(****************************************************************************************************<br>
© Syntegon Group.<br>
All rights reserved, also regarding any disposal, exploitation, reproduction, editing, distribution,<br>
as well as in the event of applications for industrial property rights.<br>
*****************************************************************************************************<br>
DESCRIPTION:<br>
A vision system's m_Configure describes housing, lens and the field of view as a frustum down to the working<br>
distance; a negative working distance gives a flat field of view at the lens.<br>
****************************************************************************************************)
METHOD PRIVATE m_VisionConfigure
VAR_INST
	fb_TempVision						: _FB_VisuVision;
	b_TempDone							: BOOL;	// the test ran
END_VAR
TEST('VisionConfigure');
IF b_TempDone THEN
	RETURN;
END_IF
b_TempDone := TRUE;

AssertTrue(Condition := fb_TempVision.m_Configure(vi_lr_FieldLength := 400, vi_lr_FieldWidth := 300,
	vi_lr_WorkingDistance := 800), Message := 'configured');
AssertEquals_UINT(Expected := 3, Actual := fb_TempVision.vo_Visu.stConfig.nBodyCount, Message := 'housing, lens, field of view');
AssertTrue(Condition := fb_TempVision.vo_Visu.stConfig.aBodies[2].eShape = E_VisuBodyShape.FRUSTUM,
	Message := 'field of view is a frustum');
AssertTrue(Condition := fb_TempVision.vo_Visu.stConfig.aBodies[2].eRole = E_VisuBodyRole.FIELD_OF_VIEW, Message := 'field of view role');
AssertEquals_LREAL(Expected := 800, Actual := fb_TempVision.vo_Visu.stConfig.aBodies[2].fHeight, Delta := 0.001,
	Message := 'field of view reaches the working distance');
AssertEquals_LREAL(Expected := -800, Actual := fb_TempVision.vo_Visu.stConfig.aBodies[2].stPose.fZ, Delta := 0.001,
	Message := 'field of view stands at the working distance below the lens');
AssertEquals_LREAL(Expected := 400, Actual := fb_TempVision.vo_Visu.stConfig.aBodies[2].fLength, Delta := 0.001,
	Message := 'field length at the bottom');

fb_TempVision.m_Configure(vi_lr_FieldLength := 400, vi_lr_FieldWidth := 300, vi_lr_WorkingDistance := -50);
AssertEquals_LREAL(Expected := 0, Actual := fb_TempVision.vo_Visu.stConfig.aBodies[2].fHeight, Delta := 0.001,
	Message := 'negative working distance: flat field of view');

TEST_FINISHED();
END_METHOD

END_FUNCTION_BLOCK

// ---- POUs/Tests/_FB_TestMachine.TcPOU
(****************************************************************************************************<br>
© Syntegon Group.<br>
All rights reserved, also regarding any disposal, exploitation, reproduction, editing, distribution,<br>
as well as in the event of applications for industrial property rights.<br>
*****************************************************************************************************<br>
DESCRIPTION:<br>
TcUnit test suite of _FB_VisuMachine: run state and simulation mode in the machine entry, machine messages set<br>
by their level, gone messages kept, and a full register making room with its oldest gone message.<br>
*****************************************************************************************************<br>
VERSION         ¦ DATE       ¦ NAME      ¦ CHANGE<br>
Syn_Visu 9.7.0  ¦ 2026-11-13 ¦ J.Willner ¦ Unit tests of the machine entry (protocol 22)<br>
****************************************************************************************************)
FUNCTION_BLOCK _FB_TestMachine EXTENDS TcUnit.FB_TestSuite
VAR
END_VAR

m_RunStateAndSimulation();
m_MessageRaisedAndCleared();
m_MessageIdZeroRefused();
m_FullRegisterMakesRoom();

(****************************************************************************************************<br>
© Syntegon Group.<br>
All rights reserved, also regarding any disposal, exploitation, reproduction, editing, distribution,<br>
as well as in the event of applications for industrial property rights.<br>
*****************************************************************************************************<br>
DESCRIPTION:<br>
A register full of active messages refuses a new one. Once some are gone, a new message takes the place of the<br>
oldest gone one (by its time): the others keep their order, the new one is last.<br>
****************************************************************************************************)
METHOD PRIVATE m_FullRegisterMakesRoom
VAR_INST
	fb_TempMachine						: _FB_VisuMachine;
	TempMachine							: ST_VisuMachine;
	b_TempDone							: BOOL;	// the test ran
END_VAR
VAR
	un_TempIndex						: UINT;
END_VAR
TEST('FullRegisterMakesRoom');
IF b_TempDone THEN
	RETURN;
END_IF
b_TempDone := TRUE;

fb_TempMachine.m_Register(vio_Machine := TempMachine);
FOR un_TempIndex := 1 TO VISU_GlobalConst_Param.VISU_un_MAX_MACHINE_MESSAGES DO
	fb_TempMachine.m_SetMessage(vi_udn_Id := un_TempIndex, vi_b_Active := TRUE,
		vi_e_Severity := E_VisuMessageSeverity.INFO, vi_str_Text := '', vi_udn_ComponentId := 0);
END_FOR
AssertEquals_UINT(Expected := VISU_GlobalConst_Param.VISU_un_MAX_MACHINE_MESSAGES, Actual := TempMachine.nMessageCount,
	Message := 'register full');
AssertFalse(Condition := fb_TempMachine.m_SetMessage(vi_udn_Id := 100, vi_b_Active := TRUE,
	vi_e_Severity := E_VisuMessageSeverity.INFO, vi_str_Text := '', vi_udn_ComponentId := 0),
	Message := 'full of active messages: a new one is refused');

(* Messages 3 and 5 go; 5 appeared earlier, so it is the oldest gone one. *)
fb_TempMachine.m_SetMessage(vi_udn_Id := 3, vi_b_Active := FALSE, vi_e_Severity := E_VisuMessageSeverity.INFO,
	vi_str_Text := '', vi_udn_ComponentId := 0);
fb_TempMachine.m_SetMessage(vi_udn_Id := 5, vi_b_Active := FALSE, vi_e_Severity := E_VisuMessageSeverity.INFO,
	vi_str_Text := '', vi_udn_ComponentId := 0);
TempMachine.aMessages[2].nTime := 2000;
TempMachine.aMessages[4].nTime := 1000;
AssertTrue(Condition := fb_TempMachine.m_SetMessage(vi_udn_Id := 100, vi_b_Active := TRUE,
	vi_e_Severity := E_VisuMessageSeverity.ERROR, vi_str_Text := 'New', vi_udn_ComponentId := 0),
	Message := 'with gone messages: a new one is listed');
AssertEquals_UINT(Expected := VISU_GlobalConst_Param.VISU_un_MAX_MACHINE_MESSAGES, Actual := TempMachine.nMessageCount,
	Message := 'still full');
AssertEquals_UDINT(Expected := 4, Actual := TempMachine.aMessages[3].nId, Message := 'message 4 before the gap');
AssertEquals_UDINT(Expected := 6, Actual := TempMachine.aMessages[4].nId, Message := 'message 5 left, 6 moved up');
AssertEquals_UDINT(Expected := 3, Actual := TempMachine.aMessages[2].nId, Message := 'message 3, gone later, stays');
AssertEquals_UDINT(Expected := 100, Actual := TempMachine.aMessages[VISU_GlobalConst_Param.VISU_un_MAX_MACHINE_MESSAGES - 1].nId,
	Message := 'the new message is last');
AssertTrue(Condition := TempMachine.aMessages[VISU_GlobalConst_Param.VISU_un_MAX_MACHINE_MESSAGES - 1].bActive,
	Message := 'the new message is active');

TEST_FINISHED();
END_METHOD

(****************************************************************************************************<br>
© Syntegon Group.<br>
All rights reserved, also regarding any disposal, exploitation, reproduction, editing, distribution,<br>
as well as in the event of applications for industrial property rights.<br>
*****************************************************************************************************<br>
DESCRIPTION:<br>
A message with id 0 is refused and not listed.<br>
****************************************************************************************************)
METHOD PRIVATE m_MessageIdZeroRefused
VAR_INST
	fb_TempMachine						: _FB_VisuMachine;
	TempMachine							: ST_VisuMachine;
	b_TempDone							: BOOL;	// the test ran
END_VAR
TEST('MessageIdZeroRefused');
IF b_TempDone THEN
	RETURN;
END_IF
b_TempDone := TRUE;

fb_TempMachine.m_Register(vio_Machine := TempMachine);
AssertFalse(Condition := fb_TempMachine.m_SetMessage(vi_udn_Id := 0, vi_b_Active := TRUE,
	vi_e_Severity := E_VisuMessageSeverity.ERROR, vi_str_Text := 'x', vi_udn_ComponentId := 0),
	Message := 'id 0 refused');
AssertEquals_UINT(Expected := 0, Actual := TempMachine.nMessageCount, Message := 'nothing listed');

TEST_FINISHED();
END_METHOD

(****************************************************************************************************<br>
© Syntegon Group.<br>
All rights reserved, also regarding any disposal, exploitation, reproduction, editing, distribution,<br>
as well as in the event of applications for industrial property rights.<br>
*****************************************************************************************************<br>
DESCRIPTION:<br>
A message set active is listed with its severity, text and component; set again it stays one entry and follows<br>
the inputs. Cleared it is gone but still listed; set active again it is the same entry, active once more. Clearing<br>
a message that was never listed lists nothing.<br>
****************************************************************************************************)
METHOD PRIVATE m_MessageRaisedAndCleared
VAR_INST
	fb_TempMachine						: _FB_VisuMachine;
	TempMachine							: ST_VisuMachine;
	b_TempDone							: BOOL;	// the test ran
END_VAR
TEST('MessageRaisedAndCleared');
IF b_TempDone THEN
	RETURN;
END_IF
b_TempDone := TRUE;

fb_TempMachine.m_Register(vio_Machine := TempMachine);
AssertTrue(Condition := fb_TempMachine.m_SetMessage(vi_udn_Id := 7, vi_b_Active := TRUE,
	vi_e_Severity := E_VisuMessageSeverity.WARNING, vi_str_Text := 'Reject bin almost full', vi_udn_ComponentId := 60),
	Message := 'a new message is listed');
AssertEquals_UINT(Expected := 1, Actual := TempMachine.nMessageCount, Message := 'one message');
AssertEquals_UDINT(Expected := 7, Actual := TempMachine.aMessages[0].nId, Message := 'its id');
AssertTrue(Condition := TempMachine.aMessages[0].bActive, Message := 'active');
AssertTrue(Condition := TempMachine.aMessages[0].eSeverity = E_VisuMessageSeverity.WARNING, Message := 'severity WARNING');
AssertEquals_STRING(Expected := 'Reject bin almost full', Actual := TempMachine.aMessages[0].sText, Message := 'its text');
AssertEquals_UDINT(Expected := 60, Actual := TempMachine.aMessages[0].nComponentId, Message := 'its component');

fb_TempMachine.m_SetMessage(vi_udn_Id := 7, vi_b_Active := TRUE, vi_e_Severity := E_VisuMessageSeverity.ERROR,
	vi_str_Text := 'Reject bin full', vi_udn_ComponentId := 60);
AssertEquals_UINT(Expected := 1, Actual := TempMachine.nMessageCount, Message := 'set again: still one message');
AssertTrue(Condition := TempMachine.aMessages[0].eSeverity = E_VisuMessageSeverity.ERROR, Message := 'severity follows');
AssertEquals_STRING(Expected := 'Reject bin full', Actual := TempMachine.aMessages[0].sText, Message := 'text follows');

fb_TempMachine.m_SetMessage(vi_udn_Id := 7, vi_b_Active := FALSE, vi_e_Severity := E_VisuMessageSeverity.ERROR,
	vi_str_Text := 'Reject bin full', vi_udn_ComponentId := 60);
AssertEquals_UINT(Expected := 1, Actual := TempMachine.nMessageCount, Message := 'cleared: still listed');
AssertFalse(Condition := TempMachine.aMessages[0].bActive, Message := 'cleared: gone');

fb_TempMachine.m_SetMessage(vi_udn_Id := 7, vi_b_Active := TRUE, vi_e_Severity := E_VisuMessageSeverity.ERROR,
	vi_str_Text := 'Reject bin full', vi_udn_ComponentId := 60);
AssertEquals_UINT(Expected := 1, Actual := TempMachine.nMessageCount, Message := 'raised again: the same entry');
AssertTrue(Condition := TempMachine.aMessages[0].bActive, Message := 'raised again: active');

AssertTrue(Condition := fb_TempMachine.m_SetMessage(vi_udn_Id := 8, vi_b_Active := FALSE,
	vi_e_Severity := E_VisuMessageSeverity.INFO, vi_str_Text := '', vi_udn_ComponentId := 0),
	Message := 'clearing an unlisted message succeeds');
AssertEquals_UINT(Expected := 1, Actual := TempMachine.nMessageCount, Message := '... and lists nothing');

TEST_FINISHED();
END_METHOD

(****************************************************************************************************<br>
© Syntegon Group.<br>
All rights reserved, also regarding any disposal, exploitation, reproduction, editing, distribution,<br>
as well as in the event of applications for industrial property rights.<br>
*****************************************************************************************************<br>
DESCRIPTION:<br>
Before m_Register the methods write nothing; after it the run state, its text and simulation mode are in the<br>
machine entry.<br>
****************************************************************************************************)
METHOD PRIVATE m_RunStateAndSimulation
VAR_INST
	fb_TempMachine						: _FB_VisuMachine;
	TempMachine							: ST_VisuMachine;
	b_TempDone							: BOOL;	// the test ran
END_VAR
TEST('RunStateAndSimulation');
IF b_TempDone THEN
	RETURN;
END_IF
b_TempDone := TRUE;

AssertFalse(Condition := fb_TempMachine.m_SetRunState(vi_e_RunState := E_VisuRunState.RUNNING, vi_str_Text := ''),
	Message := 'm_SetRunState before m_Register: FALSE');
AssertFalse(Condition := fb_TempMachine.m_SetMessage(vi_udn_Id := 1, vi_b_Active := TRUE,
	vi_e_Severity := E_VisuMessageSeverity.ERROR, vi_str_Text := 'x', vi_udn_ComponentId := 0),
	Message := 'm_SetMessage before m_Register: FALSE');

AssertTrue(Condition := fb_TempMachine.m_Register(vio_Machine := TempMachine), Message := 'm_Register');
AssertTrue(Condition := fb_TempMachine.m_SetRunState(vi_e_RunState := E_VisuRunState.FAULT, vi_str_Text := 'Vacuum lost'),
	Message := 'm_SetRunState after m_Register');
AssertTrue(Condition := fb_TempMachine.m_SetSimulation(vi_b_Simulation := TRUE), Message := 'm_SetSimulation');
AssertTrue(Condition := TempMachine.eRunState = E_VisuRunState.FAULT, Message := 'run state FAULT');
AssertEquals_STRING(Expected := 'Vacuum lost', Actual := TempMachine.sRunStateText, Message := 'run state text');
AssertTrue(Condition := TempMachine.bSimulation, Message := 'simulation mode');
AssertEquals_UINT(Expected := 0, Actual := TempMachine.nMessageCount, Message := 'no messages');

TEST_FINISHED();
END_METHOD

END_FUNCTION_BLOCK

// ---- POUs/Tests/_FB_TestConfigComponent.TcPOU
(****************************************************************************************************<br>
© Syntegon Group.<br>
All rights reserved, also regarding any disposal, exploitation, reproduction, editing, distribution,<br>
as well as in the event of applications for industrial property rights.<br>
*****************************************************************************************************<br>
DESCRIPTION:<br>
TcUnit test suite of SynConfig._FB_ConfigComponent: registration in the config manifest (m_Register, m_Id), the<br>
symbol path of vo_Config taken from the instance path, and the protocol and library version reported to the<br>
gateway.<br>
*****************************************************************************************************<br>
VERSION         ¦ DATE       ¦ NAME      ¦ CHANGE<br>
Syn_Config 2.0.0 ¦ 2026-11-11 ¦ J.Willner ¦ Unit tests<br>
****************************************************************************************************)
FUNCTION_BLOCK _FB_TestConfigComponent EXTENDS TcUnit.FB_TestSuite
VAR
	fb_PathConveyorParam				: SynConfig._FB_ConfigConveyor;	// declared here so that its instance path is known
END_VAR

m_RegisterAddsEntry();
m_RegisterIsIdempotent();
m_RegisterRejectsIdZero();
m_RegisterRejectsUsedId();
m_RegisterRejectsFullManifest();
m_RegisterSymbolPath();
m_VersionMatchesConstant();

(****************************************************************************************************<br>
© Syntegon Group.<br>
All rights reserved, also regarding any disposal, exploitation, reproduction, editing, distribution,<br>
as well as in the event of applications for industrial property rights.<br>
*****************************************************************************************************<br>
DESCRIPTION:<br>
m_Register adds an entry with the id and type of the parametrised component, gives the id through m_Id and<br>
reports the running library's protocol and library version in the manifest.<br>
****************************************************************************************************)
METHOD PRIVATE m_RegisterAddsEntry
VAR_INST
	fb_TempParam						: SynConfig._FB_ConfigDelta;
	TempManifest						: SynConfig.ST_ConfigManifest;
	b_TempDone							: BOOL;	// the test ran
END_VAR
TEST('ConfigRegisterAddsEntry');
IF b_TempDone THEN
	RETURN;
END_IF
b_TempDone := TRUE;

AssertEquals_UDINT(Expected := 0, Actual := fb_TempParam.m_Id(), Message := 'not registered: id 0');
AssertTrue(Condition := fb_TempParam.m_Register(vio_Manifest := TempManifest, vi_udn_Id := 10), Message := 'registered');
AssertEquals_UINT(Expected := 1, Actual := TempManifest.nCount, Message := 'one entry');
AssertEquals_UDINT(Expected := 10, Actual := TempManifest.aEntries[0].nId, Message := 'entry has the component id');
AssertTrue(Condition := TempManifest.aEntries[0].eType = E_VisuComponentType.DELTA, Message := 'entry has the component type');
AssertEquals_UDINT(Expected := 10, Actual := fb_TempParam.m_Id(), Message := 'm_Id gives the id');
AssertEquals_UINT(Expected := SynConfig.CONFIG_GlobalConst.CONFIG_un_PROTOCOL_VERSION, Actual := TempManifest.nProtocolVersion,
	Message := 'config protocol version reported');
AssertEquals_STRING(Expected := SynConfig.CONFIG_GlobalConst.CONFIG_str_LIBRARY_VERSION, Actual := TempManifest.sLibraryVersion,
	Message := 'library version reported');

TEST_FINISHED();
END_METHOD

(****************************************************************************************************<br>
© Syntegon Group.<br>
All rights reserved, also regarding any disposal, exploitation, reproduction, editing, distribution,<br>
as well as in the event of applications for industrial property rights.<br>
*****************************************************************************************************<br>
DESCRIPTION:<br>
m_Register is called every cycle: registering again with the same id succeeds without a second entry.<br>
****************************************************************************************************)
METHOD PRIVATE m_RegisterIsIdempotent
VAR_INST
	fb_TempParam						: SynConfig._FB_ConfigConveyor;
	TempManifest						: SynConfig.ST_ConfigManifest;
	b_TempDone							: BOOL;	// the test ran
END_VAR
TEST('ConfigRegisterIsIdempotent');
IF b_TempDone THEN
	RETURN;
END_IF
b_TempDone := TRUE;

AssertTrue(Condition := fb_TempParam.m_Register(vio_Manifest := TempManifest, vi_udn_Id := 1), Message := 'first call');
AssertTrue(Condition := fb_TempParam.m_Register(vio_Manifest := TempManifest, vi_udn_Id := 1), Message := 'second call');
AssertEquals_UINT(Expected := 1, Actual := TempManifest.nCount, Message := 'still one entry');

TEST_FINISHED();
END_METHOD

(****************************************************************************************************<br>
© Syntegon Group.<br>
All rights reserved, also regarding any disposal, exploitation, reproduction, editing, distribution,<br>
as well as in the event of applications for industrial property rights.<br>
*****************************************************************************************************<br>
DESCRIPTION:<br>
The config manifest takes CONFIG_un_MAX_MANIFEST_ENTRIES entries; a new id beyond them is refused.<br>
****************************************************************************************************)
METHOD PRIVATE m_RegisterRejectsFullManifest
VAR_INST
	fb_TempParam						: SynConfig._FB_ConfigConveyor;
	TempManifest						: SynConfig.ST_ConfigManifest;
	b_TempDone							: BOOL;	// the test ran
END_VAR
VAR
	un_TempEntry						: UINT;
END_VAR
TEST('ConfigRegisterRejectsFullManifest');
IF b_TempDone THEN
	RETURN;
END_IF
b_TempDone := TRUE;

(* Other parameter FBs have filled the manifest. *)
FOR un_TempEntry := 0 TO SynConfig.CONFIG_GlobalConst_Param.CONFIG_un_MAX_MANIFEST_ENTRIES - 1 DO
	TempManifest.aEntries[un_TempEntry].nId := UINT_TO_UDINT(un_TempEntry + 1);
	TempManifest.aEntries[un_TempEntry].eType := E_VisuComponentType.CONVEYOR;
	TempManifest.aEntries[un_TempEntry].sPath := 'P_Line.fb_Param.vo_Config';
END_FOR
TempManifest.nCount := SynConfig.CONFIG_GlobalConst_Param.CONFIG_un_MAX_MANIFEST_ENTRIES;

AssertFalse(Condition := fb_TempParam.m_Register(vio_Manifest := TempManifest, vi_udn_Id := 999), Message := 'full manifest refuses');
AssertEquals_UINT(Expected := SynConfig.CONFIG_GlobalConst_Param.CONFIG_un_MAX_MANIFEST_ENTRIES, Actual := TempManifest.nCount,
	Message := 'entry count at the limit');

TEST_FINISHED();
END_METHOD

(****************************************************************************************************<br>
© Syntegon Group.<br>
All rights reserved, also regarding any disposal, exploitation, reproduction, editing, distribution,<br>
as well as in the event of applications for industrial property rights.<br>
*****************************************************************************************************<br>
DESCRIPTION:<br>
Id 0 is no component (an unregistered Syn_Visu FB's m_Id): m_Register refuses it and adds nothing.<br>
****************************************************************************************************)
METHOD PRIVATE m_RegisterRejectsIdZero
VAR_INST
	fb_TempParam						: SynConfig._FB_ConfigConveyor;
	TempManifest						: SynConfig.ST_ConfigManifest;
	b_TempDone							: BOOL;	// the test ran
END_VAR
TEST('ConfigRegisterRejectsIdZero');
IF b_TempDone THEN
	RETURN;
END_IF
b_TempDone := TRUE;

AssertFalse(Condition := fb_TempParam.m_Register(vio_Manifest := TempManifest, vi_udn_Id := 0), Message := 'id 0 refused');
AssertEquals_UINT(Expected := 0, Actual := TempManifest.nCount, Message := 'no entry');
AssertEquals_UDINT(Expected := 0, Actual := fb_TempParam.m_Id(), Message := 'still not registered');

TEST_FINISHED();
END_METHOD

(****************************************************************************************************<br>
© Syntegon Group.<br>
All rights reserved, also regarding any disposal, exploitation, reproduction, editing, distribution,<br>
as well as in the event of applications for industrial property rights.<br>
*****************************************************************************************************<br>
DESCRIPTION:<br>
One parameter FB per component: an id already registered by another FB is refused, whether that FB has another<br>
type or the same type at another symbol path.<br>
****************************************************************************************************)
METHOD PRIVATE m_RegisterRejectsUsedId
VAR_INST
	fb_TempConveyorParam				: SynConfig._FB_ConfigConveyor;
	fb_TempOtherConveyorParam			: SynConfig._FB_ConfigConveyor;
	fb_TempDeltaParam					: SynConfig._FB_ConfigDelta;
	TempManifest						: SynConfig.ST_ConfigManifest;
	b_TempDone							: BOOL;	// the test ran
END_VAR
TEST('ConfigRegisterRejectsUsedId');
IF b_TempDone THEN
	RETURN;
END_IF
b_TempDone := TRUE;

AssertTrue(Condition := fb_TempConveyorParam.m_Register(vio_Manifest := TempManifest, vi_udn_Id := 3), Message := 'first FB registered');
AssertFalse(Condition := fb_TempDeltaParam.m_Register(vio_Manifest := TempManifest, vi_udn_Id := 3),
	Message := 'another type with the same id refused');
AssertFalse(Condition := fb_TempOtherConveyorParam.m_Register(vio_Manifest := TempManifest, vi_udn_Id := 3),
	Message := 'the same type at another path refused');
AssertEquals_UINT(Expected := 1, Actual := TempManifest.nCount, Message := 'still one entry');
AssertEquals_UDINT(Expected := 0, Actual := fb_TempDeltaParam.m_Id(), Message := 'refused FB not registered');

TEST_FINISHED();
END_METHOD

(****************************************************************************************************<br>
© Syntegon Group.<br>
All rights reserved, also regarding any disposal, exploitation, reproduction, editing, distribution,<br>
as well as in the event of applications for industrial property rights.<br>
*****************************************************************************************************<br>
DESCRIPTION:<br>
The manifest entry's symbol path is the instance path without TwinCAT project and PLC project, plus<br>
'.vo_Config': the path the gateway reads and writes over ADS.<br>
****************************************************************************************************)
METHOD PRIVATE m_RegisterSymbolPath
VAR_INST
	TempManifest						: SynConfig.ST_ConfigManifest;
	b_TempDone							: BOOL;	// the test ran
END_VAR
TEST('ConfigRegisterSymbolPath');
IF b_TempDone THEN
	RETURN;
END_IF
b_TempDone := TRUE;

fb_PathConveyorParam.m_Register(vio_Manifest := TempManifest, vi_udn_Id := 1);
AssertEquals_STRING(Expected := 'P_TestRun.fb_TestConfigComponent.fb_PathConveyorParam.vo_Config',
	Actual := TempManifest.aEntries[0].sPath, Message := 'symbol path of vo_Config without TwinCAT and PLC project');

TEST_FINISHED();
END_METHOD

(****************************************************************************************************<br>
© Syntegon Group.<br>
All rights reserved, also regarding any disposal, exploitation, reproduction, editing, distribution,<br>
as well as in the event of applications for industrial property rights.<br>
*****************************************************************************************************<br>
DESCRIPTION:<br>
_FC_GetVersionSynConfig and CONFIG_str_LIBRARY_VERSION name the same version: both are bumped together.<br>
****************************************************************************************************)
METHOD PRIVATE m_VersionMatchesConstant
VAR_INST
	b_TempDone							: BOOL;	// the test ran
END_VAR
VAR
	str_TempVersion						: STRING(31);	// major.minor.revision from _FC_GetVersionSynConfig
END_VAR
TEST('ConfigVersionMatchesConstant');
IF b_TempDone THEN
	RETURN;
END_IF
b_TempDone := TRUE;

str_TempVersion := CONCAT(UINT_TO_STRING(SynConfig._FC_GetVersionSynConfig(vi_n_VersionElement := 1)), '.');
str_TempVersion := CONCAT(str_TempVersion, UINT_TO_STRING(SynConfig._FC_GetVersionSynConfig(vi_n_VersionElement := 2)));
str_TempVersion := CONCAT(str_TempVersion, '.');
str_TempVersion := CONCAT(str_TempVersion, UINT_TO_STRING(SynConfig._FC_GetVersionSynConfig(vi_n_VersionElement := 3)));
AssertEquals_STRING(Expected := SynConfig.CONFIG_GlobalConst.CONFIG_str_LIBRARY_VERSION, Actual := str_TempVersion,
	Message := '_FC_GetVersionSynConfig matches CONFIG_str_LIBRARY_VERSION');
AssertEquals_UINT(Expected := 16#FFFF, Actual := SynConfig._FC_GetVersionSynConfig(vi_n_VersionElement := 4),
	Message := 'unknown version element gives 16#FFFF');

TEST_FINISHED();
END_METHOD

END_FUNCTION_BLOCK

// ---- POUs/Tests/_FB_TestConfigStaging.TcPOU
(****************************************************************************************************<br>
© Syntegon Group.<br>
All rights reserved, also regarding any disposal, exploitation, reproduction, editing, distribution,<br>
as well as in the event of applications for industrial property rights.<br>
*****************************************************************************************************<br>
DESCRIPTION:<br>
TcUnit test suite of a parameter FB's m_Cycle (ADR 0017), on SynConfig._FB_ConfigConveyor: the program values<br>
while no set is active, a staged set taken over, waiting while the application does not allow it, rejected on<br>
another active version or when invalid, and a reset back to the program values. The tests write vo_Config's<br>
stStaging and stStaged as the gateway does over ADS.<br>
*****************************************************************************************************<br>
VERSION         ¦ DATE       ¦ NAME      ¦ CHANGE<br>
Syn_Config 2.0.0 ¦ 2026-11-11 ¦ J.Willner ¦ Unit tests<br>
Syn_Config 2.3.0 ¦ 2026-11-14 ¦ J.Willner ¦ The lifecycle of every parameter FB type<br>
****************************************************************************************************)
FUNCTION_BLOCK _FB_TestConfigStaging EXTENDS TcUnit.FB_TestSuite

m_ProgramValuesWithoutSet();
m_StagedSetTakenOver();
m_StagedSetWaitsUntilAllowed();
m_StagedSetOnOtherVersionRejected();
m_ResetReturnsToProgramValues();
m_InvalidProductTypesRejected();
m_EveryTypeRunsTheLifecycle();

(****************************************************************************************************<br>
© Syntegon Group.<br>
All rights reserved, also regarding any disposal, exploitation, reproduction, editing, distribution,<br>
as well as in the event of applications for industrial property rights.<br>
*****************************************************************************************************<br>
DESCRIPTION:<br>
Every parameter FB type runs the same staging lifecycle as the conveyor: a set staged on version 0 is taken over<br>
as version 1, a set staged on version 0 again is rejected (version 1 is active), and a reset returns to the<br>
program values under version 0. The machine FB's recipe has its own suite (_FB_TestConfigMachine).<br>
****************************************************************************************************)
METHOD PRIVATE m_EveryTypeRunsTheLifecycle
VAR_INST
	fb_TempDelta						: SynConfig._FB_ConfigDelta;
	TempDeltaDefault					: SynConfig.ST_ConfigDeltaParam;
	TempDeltaStaged						: SynConfig.ST_ConfigDeltaParam;
	TempDeltaSet						: SynConfig.ST_ConfigDeltaSet;
	fb_TempGantry						: SynConfig._FB_ConfigXtsGantry;
	TempGantryDefault					: SynConfig.ST_ConfigXtsGantryParam;
	TempGantryStaged					: SynConfig.ST_ConfigXtsGantryParam;
	TempGantrySet						: SynConfig.ST_ConfigXtsGantrySet;
	fb_TempLoop							: SynConfig._FB_ConfigXtsLoop;
	TempLoopDefault						: SynConfig.ST_ConfigXtsLoopParam;
	TempLoopStaged						: SynConfig.ST_ConfigXtsLoopParam;
	TempLoopSet							: SynConfig.ST_ConfigXtsLoopSet;
	fb_TempCartesian					: SynConfig._FB_ConfigCartesian;
	TempCartesianDefault				: SynConfig.ST_ConfigCartesianParam;
	TempCartesianStaged					: SynConfig.ST_ConfigCartesianParam;
	TempCartesianSet					: SynConfig.ST_ConfigCartesianSet;
	fb_TempVision						: SynConfig._FB_ConfigVision;
	TempVisionDefault					: SynConfig.ST_ConfigBodyComponentParam;
	TempVisionStaged					: SynConfig.ST_ConfigBodyComponentParam;
	TempVisionSet						: SynConfig.ST_ConfigBodyComponentSet;
	b_TempDone							: BOOL;	// the test ran
END_VAR
VAR
	b_TempChanged						: ARRAY[1..5, 1..3] OF BOOL;	// per type and step: m_Cycle's result
	e_TempResult						: ARRAY[1..5, 1..3] OF SynConfig.E_ConfigResult;	// per type and step: stStatus.eResult
	udn_TempVersion						: ARRAY[1..5, 1..3] OF UDINT;	// [-] per type and step: stStatus.nActiveVersion
	lr_TempX							: ARRAY[1..5, 1..3] OF LREAL;	// [mm] per type and step: X of the effective pose
	TempPose							: ST_VisuPose;
	un_TempStep							: UINT;	// [-] 1 = take-over, 2 = stale version, 3 = reset
	un_TempType							: UINT;
	p_TempDelta							: POINTER TO SynConfig.ST_ConfigDeltaParam;
	p_TempGantry						: POINTER TO SynConfig.ST_ConfigXtsGantryParam;
	p_TempLoop							: POINTER TO SynConfig.ST_ConfigXtsLoopParam;
	p_TempCartesian						: POINTER TO SynConfig.ST_ConfigCartesianParam;
	p_TempVision						: POINTER TO SynConfig.ST_ConfigBodyComponentParam;
END_VAR
VAR CONSTANT
	str_TYPE_NAMES						: ARRAY[1..5] OF STRING(20) := ['Delta', 'XTS gantry', 'XTS loop', 'Cartesian', 'Vision'];
END_VAR
TEST('ConfigEveryTypeRunsTheLifecycle');
IF b_TempDone THEN
	RETURN;
END_IF
b_TempDone := TRUE;


(****************************************************************************************************
THREE STEPS PER TYPE: TAKE-OVER, STALE VERSION, RESET
****************************************************************************************************)
(* Delta *)
TempDeltaDefault.stPose.fX := 100;
TempDeltaStaged.stPose.fX := 250;
p_TempDelta := ADR(fb_TempDelta.vo_Config.stStaged);
FOR un_TempStep := 1 TO 3 DO
	p_TempDelta^ := TempDeltaStaged;
	_FC_TestConfigStage(vi_p_Staging := ADR(fb_TempDelta.vo_Config.stStaging), vi_udn_BaseVersion := 0,
		vi_udn_StageId := UINT_TO_UDINT(un_TempStep), vi_b_Reset := un_TempStep = 3);
	b_TempChanged[1, un_TempStep] := fb_TempDelta.m_Cycle(vio_Default := TempDeltaDefault, vio_Set := TempDeltaSet,
		vi_b_ApplyAllowed := TRUE);
	e_TempResult[1, un_TempStep] := fb_TempDelta.vo_Config.stStatus.eResult;
	udn_TempVersion[1, un_TempStep] := fb_TempDelta.vo_Config.stStatus.nActiveVersion;
	TempPose := fb_TempDelta.m_Pose();
	lr_TempX[1, un_TempStep] := TempPose.fX;
END_FOR

(* XTS gantry: a track needs a module *)
TempGantryDefault.stPose.fX := 100;
TempGantryStaged.stPose.fX := 250;
TempGantryStaged.nModuleCount := 1;
TempGantryStaged.aModules[0].fLength := 250;
p_TempGantry := ADR(fb_TempGantry.vo_Config.stStaged);
FOR un_TempStep := 1 TO 3 DO
	p_TempGantry^ := TempGantryStaged;
	_FC_TestConfigStage(vi_p_Staging := ADR(fb_TempGantry.vo_Config.stStaging), vi_udn_BaseVersion := 0,
		vi_udn_StageId := UINT_TO_UDINT(un_TempStep), vi_b_Reset := un_TempStep = 3);
	b_TempChanged[2, un_TempStep] := fb_TempGantry.m_Cycle(vio_Default := TempGantryDefault, vio_Set := TempGantrySet,
		vi_b_ApplyAllowed := TRUE);
	e_TempResult[2, un_TempStep] := fb_TempGantry.vo_Config.stStatus.eResult;
	udn_TempVersion[2, un_TempStep] := fb_TempGantry.vo_Config.stStatus.nActiveVersion;
	TempPose := fb_TempGantry.m_Pose();
	lr_TempX[2, un_TempStep] := TempPose.fX;
END_FOR

(* XTS loop: a track needs a module *)
TempLoopDefault.stPose.fX := 100;
TempLoopStaged.stPose.fX := 250;
TempLoopStaged.nModuleCount := 1;
TempLoopStaged.aModules[0].fLength := 250;
p_TempLoop := ADR(fb_TempLoop.vo_Config.stStaged);
FOR un_TempStep := 1 TO 3 DO
	p_TempLoop^ := TempLoopStaged;
	_FC_TestConfigStage(vi_p_Staging := ADR(fb_TempLoop.vo_Config.stStaging), vi_udn_BaseVersion := 0,
		vi_udn_StageId := UINT_TO_UDINT(un_TempStep), vi_b_Reset := un_TempStep = 3);
	b_TempChanged[3, un_TempStep] := fb_TempLoop.m_Cycle(vio_Default := TempLoopDefault, vio_Set := TempLoopSet,
		vi_b_ApplyAllowed := TRUE);
	e_TempResult[3, un_TempStep] := fb_TempLoop.vo_Config.stStatus.eResult;
	udn_TempVersion[3, un_TempStep] := fb_TempLoop.vo_Config.stStatus.nActiveVersion;
	TempPose := fb_TempLoop.m_Pose();
	lr_TempX[3, un_TempStep] := TempPose.fX;
END_FOR

(* Cartesian *)
TempCartesianDefault.stPose.fX := 100;
TempCartesianStaged.stPose.fX := 250;
p_TempCartesian := ADR(fb_TempCartesian.vo_Config.stStaged);
FOR un_TempStep := 1 TO 3 DO
	p_TempCartesian^ := TempCartesianStaged;
	_FC_TestConfigStage(vi_p_Staging := ADR(fb_TempCartesian.vo_Config.stStaging), vi_udn_BaseVersion := 0,
		vi_udn_StageId := UINT_TO_UDINT(un_TempStep), vi_b_Reset := un_TempStep = 3);
	b_TempChanged[4, un_TempStep] := fb_TempCartesian.m_Cycle(vio_Default := TempCartesianDefault,
		vio_Set := TempCartesianSet, vi_b_ApplyAllowed := TRUE);
	e_TempResult[4, un_TempStep] := fb_TempCartesian.vo_Config.stStatus.eResult;
	udn_TempVersion[4, un_TempStep] := fb_TempCartesian.vo_Config.stStatus.nActiveVersion;
	TempPose := fb_TempCartesian.m_Pose();
	lr_TempX[4, un_TempStep] := TempPose.fX;
END_FOR

(* Vision system, for the body components *)
TempVisionDefault.stPose.fX := 100;
TempVisionStaged.stPose.fX := 250;
p_TempVision := ADR(fb_TempVision.vo_Config.stStaged);
FOR un_TempStep := 1 TO 3 DO
	p_TempVision^ := TempVisionStaged;
	_FC_TestConfigStage(vi_p_Staging := ADR(fb_TempVision.vo_Config.stStaging), vi_udn_BaseVersion := 0,
		vi_udn_StageId := UINT_TO_UDINT(un_TempStep), vi_b_Reset := un_TempStep = 3);
	b_TempChanged[5, un_TempStep] := fb_TempVision.m_Cycle(vio_Default := TempVisionDefault, vio_Set := TempVisionSet,
		vi_b_ApplyAllowed := TRUE);
	e_TempResult[5, un_TempStep] := fb_TempVision.vo_Config.stStatus.eResult;
	udn_TempVersion[5, un_TempStep] := fb_TempVision.vo_Config.stStatus.nActiveVersion;
	TempPose := fb_TempVision.m_Pose();
	lr_TempX[5, un_TempStep] := TempPose.fX;
END_FOR


(****************************************************************************************************
THE SAME RESULTS FOR EVERY TYPE
****************************************************************************************************)
FOR un_TempType := 1 TO 5 DO
	AssertTrue(Condition := b_TempChanged[un_TempType, 1], Message := CONCAT(str_TYPE_NAMES[un_TempType], ': taken over'));
	AssertEquals_UDINT(Expected := 1, Actual := udn_TempVersion[un_TempType, 1],
		Message := CONCAT(str_TYPE_NAMES[un_TempType], ': version 1 active'));
	AssertEquals_LREAL(Expected := 250, Actual := lr_TempX[un_TempType, 1], Delta := 0.001,
		Message := CONCAT(str_TYPE_NAMES[un_TempType], ': staged pose effective'));
	AssertFalse(Condition := b_TempChanged[un_TempType, 2],
		Message := CONCAT(str_TYPE_NAMES[un_TempType], ': stale version not taken over'));
	AssertTrue(Condition := e_TempResult[un_TempType, 2] = SynConfig.E_ConfigResult.REJECTED,
		Message := CONCAT(str_TYPE_NAMES[un_TempType], ': stale version rejected'));
	AssertEquals_UDINT(Expected := 1, Actual := udn_TempVersion[un_TempType, 2],
		Message := CONCAT(str_TYPE_NAMES[un_TempType], ': version 1 stays'));
	AssertTrue(Condition := b_TempChanged[un_TempType, 3], Message := CONCAT(str_TYPE_NAMES[un_TempType], ': reset'));
	AssertEquals_UDINT(Expected := 0, Actual := udn_TempVersion[un_TempType, 3],
		Message := CONCAT(str_TYPE_NAMES[un_TempType], ': version 0 after the reset'));
	AssertEquals_LREAL(Expected := 100, Actual := lr_TempX[un_TempType, 3], Delta := 0.001,
		Message := CONCAT(str_TYPE_NAMES[un_TempType], ': program pose again'));
END_FOR

TEST_FINISHED();
END_METHOD

(****************************************************************************************************<br>
© Syntegon Group.<br>
All rights reserved, also regarding any disposal, exploitation, reproduction, editing, distribution,<br>
as well as in the event of applications for industrial property rights.<br>
*****************************************************************************************************<br>
DESCRIPTION:<br>
A conveyor set is rejected with the reason when a product type has no number, a number is used twice or there<br>
are more product types than the list holds; the active set stays as it was.<br>
****************************************************************************************************)
METHOD PRIVATE m_InvalidProductTypesRejected
VAR_INST
	fb_TempParam						: SynConfig._FB_ConfigConveyor;
	TempDefault							: SynConfig.ST_ConfigConveyorParam;
	TempSet								: SynConfig.ST_ConfigConveyorSet;
	b_TempDone							: BOOL;	// the test ran
END_VAR
VAR
	TempStaged							: SynConfig.ST_ConfigConveyorParam;
END_VAR
TEST('ConfigInvalidProductTypesRejected');
IF b_TempDone THEN
	RETURN;
END_IF
b_TempDone := TRUE;

TempDefault := m_ValidSet(vi_lr_X := 100);

(* A product type without a number. *)
TempStaged := m_ValidSet(vi_lr_X := 250);
TempStaged.aProductTypes[1].nId := 0;
m_Stage(vio_Param := fb_TempParam, vio_Staged := TempStaged, vi_udn_BaseVersion := 0, vi_udn_StageId := 1);
AssertFalse(Condition := fb_TempParam.m_Cycle(vio_Default := TempDefault, vio_Set := TempSet, vi_b_ApplyAllowed := TRUE),
	Message := 'type without a number: not taken over');
AssertTrue(Condition := fb_TempParam.vo_Config.stStatus.eResult = SynConfig.E_ConfigResult.REJECTED, Message := 'rejected');
AssertEquals_STRING(Expected := 'A product type without a number', Actual := fb_TempParam.vo_Config.stStatus.sMessage,
	Message := 'reason: no number');

(* A number used twice. *)
TempStaged := m_ValidSet(vi_lr_X := 250);
TempStaged.aProductTypes[0].nId := 3;
TempStaged.aProductTypes[1].nId := 3;
m_Stage(vio_Param := fb_TempParam, vio_Staged := TempStaged, vi_udn_BaseVersion := 0, vi_udn_StageId := 2);
AssertFalse(Condition := fb_TempParam.m_Cycle(vio_Default := TempDefault, vio_Set := TempSet, vi_b_ApplyAllowed := TRUE),
	Message := 'number twice: not taken over');
AssertEquals_STRING(Expected := 'Product type 3 is defined twice', Actual := fb_TempParam.vo_Config.stStatus.sMessage,
	Message := 'reason: defined twice');

(* More product types than the list holds. *)
TempStaged := m_ValidSet(vi_lr_X := 250);
TempStaged.nProductTypeCount := VISU_GlobalConst_Param.VISU_un_MAX_PRODUCT_TYPES + 1;
m_Stage(vio_Param := fb_TempParam, vio_Staged := TempStaged, vi_udn_BaseVersion := 0, vi_udn_StageId := 3);
AssertFalse(Condition := fb_TempParam.m_Cycle(vio_Default := TempDefault, vio_Set := TempSet, vi_b_ApplyAllowed := TRUE),
	Message := 'too many types: not taken over');
AssertEquals_STRING(Expected := CONCAT('More than ', CONCAT(UINT_TO_STRING(VISU_GlobalConst_Param.VISU_un_MAX_PRODUCT_TYPES),
	' product types')), Actual := fb_TempParam.vo_Config.stStatus.sMessage, Message := 'reason: too many');
AssertEquals_UDINT(Expected := 3, Actual := fb_TempParam.vo_Config.stStatus.nHandledStageId, Message := 'last stage id handled');

AssertFalse(Condition := TempSet.bValid, Message := 'still no active set');
AssertEquals_LREAL(Expected := 100, Actual := fb_TempParam.vo_Config.stActive.stPose.fX, Delta := 0.001,
	Message := 'program values still effective');

TEST_FINISHED();
END_METHOD

(****************************************************************************************************<br>
© Syntegon Group.<br>
All rights reserved, also regarding any disposal, exploitation, reproduction, editing, distribution,<br>
as well as in the event of applications for industrial property rights.<br>
*****************************************************************************************************<br>
DESCRIPTION:<br>
Without an active set the program values are effective, under version 0, and nothing has been handled.<br>
****************************************************************************************************)
METHOD PRIVATE m_ProgramValuesWithoutSet
VAR_INST
	fb_TempParam						: SynConfig._FB_ConfigConveyor;
	TempDefault							: SynConfig.ST_ConfigConveyorParam;
	TempSet								: SynConfig.ST_ConfigConveyorSet;
	b_TempDone							: BOOL;	// the test ran
END_VAR
VAR
	TempPose							: ST_VisuPose;
END_VAR
TEST('ConfigProgramValuesWithoutSet');
IF b_TempDone THEN
	RETURN;
END_IF
b_TempDone := TRUE;

TempDefault := m_ValidSet(vi_lr_X := 100);
AssertFalse(Condition := fb_TempParam.m_Cycle(vio_Default := TempDefault, vio_Set := TempSet, vi_b_ApplyAllowed := TRUE),
	Message := 'nothing staged: no change');
TempPose := fb_TempParam.m_Pose();
AssertEquals_LREAL(Expected := 100, Actual := TempPose.fX, Delta := 0.001, Message := 'program pose effective');
AssertEquals_UINT(Expected := 2, Actual := fb_TempParam.vo_Config.stActive.nProductTypeCount, Message := 'program product types effective');
AssertEquals_UDINT(Expected := 0, Actual := fb_TempParam.vo_Config.stStatus.nActiveVersion, Message := 'version 0: program values');
AssertTrue(Condition := fb_TempParam.vo_Config.stStatus.eResult = SynConfig.E_ConfigResult.NONE, Message := 'nothing handled');

TEST_FINISHED();
END_METHOD

(****************************************************************************************************<br>
© Syntegon Group.<br>
All rights reserved, also regarding any disposal, exploitation, reproduction, editing, distribution,<br>
as well as in the event of applications for industrial property rights.<br>
*****************************************************************************************************<br>
DESCRIPTION:<br>
A reset makes the active set invalid at once (also while a take-over is not allowed): the program values apply<br>
under version 0. Versions never repeat: the next set taken over gets version 2, not 1.<br>
****************************************************************************************************)
METHOD PRIVATE m_ResetReturnsToProgramValues
VAR_INST
	fb_TempParam						: SynConfig._FB_ConfigConveyor;
	TempDefault							: SynConfig.ST_ConfigConveyorParam;
	TempSet								: SynConfig.ST_ConfigConveyorSet;
	b_TempDone							: BOOL;	// the test ran
END_VAR
VAR
	TempStaged							: SynConfig.ST_ConfigConveyorParam;
END_VAR
TEST('ConfigResetReturnsToProgramValues');
IF b_TempDone THEN
	RETURN;
END_IF
b_TempDone := TRUE;

TempDefault := m_ValidSet(vi_lr_X := 100);
TempStaged := m_ValidSet(vi_lr_X := 250);
m_Stage(vio_Param := fb_TempParam, vio_Staged := TempStaged, vi_udn_BaseVersion := 0, vi_udn_StageId := 1);
fb_TempParam.m_Cycle(vio_Default := TempDefault, vio_Set := TempSet, vi_b_ApplyAllowed := TRUE);
AssertEquals_UDINT(Expected := 1, Actual := fb_TempParam.vo_Config.stStatus.nActiveVersion, Message := 'version 1 active');

_FC_TestConfigStage(vi_p_Staging := ADR(fb_TempParam.vo_Config.stStaging), vi_udn_BaseVersion := 1, vi_udn_StageId := 2,
	vi_b_Reset := TRUE);
AssertTrue(Condition := fb_TempParam.m_Cycle(vio_Default := TempDefault, vio_Set := TempSet, vi_b_ApplyAllowed := FALSE),
	Message := 'reset handled, even while not allowed');
AssertFalse(Condition := TempSet.bValid, Message := 'active set invalid');
AssertEquals_UDINT(Expected := 0, Actual := fb_TempParam.vo_Config.stStatus.nActiveVersion, Message := 'version 0');
AssertEquals_LREAL(Expected := 100, Actual := fb_TempParam.vo_Config.stActive.stPose.fX, Delta := 0.001,
	Message := 'program values effective again');
AssertTrue(Condition := fb_TempParam.vo_Config.stStatus.eResult = SynConfig.E_ConfigResult.APPLIED, Message := 'reset applied');
AssertEquals_UDINT(Expected := 2, Actual := fb_TempParam.vo_Config.stStatus.nHandledStageId, Message := 'stage id handled');
AssertFalse(Condition := fb_TempParam.vo_Config.stStaging.bReset, Message := 'reset flag cleared');

m_Stage(vio_Param := fb_TempParam, vio_Staged := TempStaged, vi_udn_BaseVersion := 0, vi_udn_StageId := 3);
fb_TempParam.m_Cycle(vio_Default := TempDefault, vio_Set := TempSet, vi_b_ApplyAllowed := TRUE);
AssertEquals_UDINT(Expected := 2, Actual := fb_TempParam.vo_Config.stStatus.nActiveVersion, Message := 'next set gets version 2');

TEST_FINISHED();
END_METHOD

(****************************************************************************************************<br>
© Syntegon Group.<br>
All rights reserved, also regarding any disposal, exploitation, reproduction, editing, distribution,<br>
as well as in the event of applications for industrial property rights.<br>
*****************************************************************************************************<br>
DESCRIPTION:<br>
Stages a set on a conveyor's parameter FB as the gateway does: the set into vo_Config.stStaged, then stStaging<br>
(_FC_TestConfigStage). The FB handles it in its next m_Cycle.<br>
****************************************************************************************************)
METHOD PRIVATE m_Stage : BOOL
VAR_IN_OUT
	vio_Param							: SynConfig._FB_ConfigConveyor;	// the parameter FB under test
END_VAR
VAR_IN_OUT CONSTANT
	vio_Staged							: SynConfig.ST_ConfigConveyorParam;	// the set to stage
END_VAR
VAR_INPUT
	vi_udn_BaseVersion					: UDINT;	// [-] active version the set is based on
	vi_udn_StageId						: UDINT;	// [-] the gateway's id of this staging
END_VAR
VAR
	p_TempStaged						: POINTER TO SynConfig.ST_ConfigConveyorParam;
END_VAR
p_TempStaged := ADR(vio_Param.vo_Config.stStaged);
p_TempStaged^ := vio_Staged;
m_Stage := _FC_TestConfigStage(vi_p_Staging := ADR(vio_Param.vo_Config.stStaging), vi_udn_BaseVersion := vi_udn_BaseVersion,
	vi_udn_StageId := vi_udn_StageId, vi_b_Reset := FALSE);
END_METHOD

(****************************************************************************************************<br>
© Syntegon Group.<br>
All rights reserved, also regarding any disposal, exploitation, reproduction, editing, distribution,<br>
as well as in the event of applications for industrial property rights.<br>
*****************************************************************************************************<br>
DESCRIPTION:<br>
A set staged on another version than the active one is rejected with the reason, even while a take-over is<br>
allowed: someone else changed the set since the configurator read it.<br>
****************************************************************************************************)
METHOD PRIVATE m_StagedSetOnOtherVersionRejected
VAR_INST
	fb_TempParam						: SynConfig._FB_ConfigConveyor;
	TempDefault							: SynConfig.ST_ConfigConveyorParam;
	TempSet								: SynConfig.ST_ConfigConveyorSet;
	b_TempDone							: BOOL;	// the test ran
END_VAR
VAR
	TempStaged							: SynConfig.ST_ConfigConveyorParam;
END_VAR
TEST('ConfigStagedSetOnOtherVersionRejected');
IF b_TempDone THEN
	RETURN;
END_IF
b_TempDone := TRUE;

TempDefault := m_ValidSet(vi_lr_X := 100);
TempStaged := m_ValidSet(vi_lr_X := 250);
m_Stage(vio_Param := fb_TempParam, vio_Staged := TempStaged, vi_udn_BaseVersion := 5, vi_udn_StageId := 9);

AssertFalse(Condition := fb_TempParam.m_Cycle(vio_Default := TempDefault, vio_Set := TempSet, vi_b_ApplyAllowed := TRUE),
	Message := 'not taken over');
AssertTrue(Condition := fb_TempParam.vo_Config.stStatus.eResult = SynConfig.E_ConfigResult.REJECTED, Message := 'rejected');
AssertEquals_STRING(Expected := 'Based on version 5, but version 0 is active', Actual := fb_TempParam.vo_Config.stStatus.sMessage,
	Message := 'the reason');
AssertEquals_UDINT(Expected := 9, Actual := fb_TempParam.vo_Config.stStatus.nHandledStageId, Message := 'stage id handled');
AssertFalse(Condition := fb_TempParam.vo_Config.stStaging.bStaged, Message := 'staged flag cleared');
AssertFalse(Condition := TempSet.bValid, Message := 'no active set');

TEST_FINISHED();
END_METHOD

(****************************************************************************************************<br>
© Syntegon Group.<br>
All rights reserved, also regarding any disposal, exploitation, reproduction, editing, distribution,<br>
as well as in the event of applications for industrial property rights.<br>
*****************************************************************************************************<br>
DESCRIPTION:<br>
A set staged on the active version is taken over while the application allows it: it becomes the active set<br>
under version 1 and the effective values, the status names the stage id as applied and the flags are cleared.<br>
****************************************************************************************************)
METHOD PRIVATE m_StagedSetTakenOver
VAR_INST
	fb_TempParam						: SynConfig._FB_ConfigConveyor;
	TempDefault							: SynConfig.ST_ConfigConveyorParam;
	TempSet								: SynConfig.ST_ConfigConveyorSet;
	b_TempDone							: BOOL;	// the test ran
END_VAR
VAR
	TempPose							: ST_VisuPose;
	TempStaged							: SynConfig.ST_ConfigConveyorParam;
END_VAR
TEST('ConfigStagedSetTakenOver');
IF b_TempDone THEN
	RETURN;
END_IF
b_TempDone := TRUE;

TempDefault := m_ValidSet(vi_lr_X := 100);
TempStaged := m_ValidSet(vi_lr_X := 250);
m_Stage(vio_Param := fb_TempParam, vio_Staged := TempStaged, vi_udn_BaseVersion := 0, vi_udn_StageId := 7);

AssertTrue(Condition := fb_TempParam.m_Cycle(vio_Default := TempDefault, vio_Set := TempSet, vi_b_ApplyAllowed := TRUE),
	Message := 'set taken over');
AssertTrue(Condition := TempSet.bValid, Message := 'active set valid');
AssertEquals_UDINT(Expected := 1, Actual := TempSet.nVersion, Message := 'first version');
AssertEquals_UDINT(Expected := 1, Actual := fb_TempParam.vo_Config.stStatus.nActiveVersion, Message := 'status names the version');
AssertEquals_UDINT(Expected := 7, Actual := fb_TempParam.vo_Config.stStatus.nHandledStageId, Message := 'stage id handled');
AssertTrue(Condition := fb_TempParam.vo_Config.stStatus.eResult = SynConfig.E_ConfigResult.APPLIED, Message := 'applied');
AssertEquals_STRING(Expected := '', Actual := fb_TempParam.vo_Config.stStatus.sMessage, Message := 'no message');
AssertFalse(Condition := fb_TempParam.vo_Config.stStaging.bStaged, Message := 'staged flag cleared');
TempPose := fb_TempParam.m_Pose();
AssertEquals_LREAL(Expected := 250, Actual := TempPose.fX, Delta := 0.001, Message := 'staged pose effective');

AssertFalse(Condition := fb_TempParam.m_Cycle(vio_Default := TempDefault, vio_Set := TempSet, vi_b_ApplyAllowed := TRUE),
	Message := 'next cycle: no change');
AssertEquals_UDINT(Expected := 1, Actual := fb_TempParam.vo_Config.stStatus.nActiveVersion, Message := 'still version 1');

TEST_FINISHED();
END_METHOD

(****************************************************************************************************<br>
© Syntegon Group.<br>
All rights reserved, also regarding any disposal, exploitation, reproduction, editing, distribution,<br>
as well as in the event of applications for industrial property rights.<br>
*****************************************************************************************************<br>
DESCRIPTION:<br>
While the application does not allow a take-over the staged set waits (PENDING, still staged, the program values<br>
stay effective); it is taken over in the first cycle that allows it.<br>
****************************************************************************************************)
METHOD PRIVATE m_StagedSetWaitsUntilAllowed
VAR_INST
	fb_TempParam						: SynConfig._FB_ConfigConveyor;
	TempDefault							: SynConfig.ST_ConfigConveyorParam;
	TempSet								: SynConfig.ST_ConfigConveyorSet;
	b_TempDone							: BOOL;	// the test ran
END_VAR
VAR
	TempStaged							: SynConfig.ST_ConfigConveyorParam;
END_VAR
TEST('ConfigStagedSetWaitsUntilAllowed');
IF b_TempDone THEN
	RETURN;
END_IF
b_TempDone := TRUE;

TempDefault := m_ValidSet(vi_lr_X := 100);
TempStaged := m_ValidSet(vi_lr_X := 250);
m_Stage(vio_Param := fb_TempParam, vio_Staged := TempStaged, vi_udn_BaseVersion := 0, vi_udn_StageId := 3);

AssertFalse(Condition := fb_TempParam.m_Cycle(vio_Default := TempDefault, vio_Set := TempSet, vi_b_ApplyAllowed := FALSE),
	Message := 'not allowed: not taken over');
AssertTrue(Condition := fb_TempParam.vo_Config.stStatus.eResult = SynConfig.E_ConfigResult.PENDING, Message := 'pending');
AssertTrue(Condition := fb_TempParam.vo_Config.stStaging.bStaged, Message := 'still staged');
AssertFalse(Condition := TempSet.bValid, Message := 'no active set yet');
AssertEquals_LREAL(Expected := 100, Actual := fb_TempParam.vo_Config.stActive.stPose.fX, Delta := 0.001,
	Message := 'program values still effective');

AssertTrue(Condition := fb_TempParam.m_Cycle(vio_Default := TempDefault, vio_Set := TempSet, vi_b_ApplyAllowed := TRUE),
	Message := 'allowed: taken over');
AssertTrue(Condition := fb_TempParam.vo_Config.stStatus.eResult = SynConfig.E_ConfigResult.APPLIED, Message := 'applied');
AssertEquals_UDINT(Expected := 3, Actual := fb_TempParam.vo_Config.stStatus.nHandledStageId, Message := 'stage id handled');

TEST_FINISHED();
END_METHOD

(****************************************************************************************************<br>
© Syntegon Group.<br>
All rights reserved, also regarding any disposal, exploitation, reproduction, editing, distribution,<br>
as well as in the event of applications for industrial property rights.<br>
*****************************************************************************************************<br>
DESCRIPTION:<br>
A conveyor parameter set that can be taken over: the pose at X = vi_lr_X and two product types (1 and 2).<br>
****************************************************************************************************)
METHOD PRIVATE m_ValidSet : SynConfig.ST_ConfigConveyorParam
VAR_INPUT
	vi_lr_X								: LREAL;	// [mm] X of the pose, to tell sets apart
END_VAR
m_ValidSet.stPose.fX := vi_lr_X;
m_ValidSet.stOriginShift.fX := 50;
m_ValidSet.nProductTypeCount := 2;
m_ValidSet.aProductTypes[0].nId := 1;
m_ValidSet.aProductTypes[0].fLength := 120;
m_ValidSet.aProductTypes[0].fWidth := 80;
m_ValidSet.aProductTypes[0].fHeight := 40;
m_ValidSet.aProductTypes[0].eShape := E_VisuProductShape.BOX;
m_ValidSet.aProductTypes[1].nId := 2;
m_ValidSet.aProductTypes[1].fLength := 66;
m_ValidSet.aProductTypes[1].fWidth := 66;
m_ValidSet.aProductTypes[1].fHeight := 120;
m_ValidSet.aProductTypes[1].eShape := E_VisuProductShape.CYLINDER;
END_METHOD

END_FUNCTION_BLOCK

// ---- POUs/Tests/_FC_TestConfigStage.TcPOU
(****************************************************************************************************<br>
© Syntegon Group.<br>
All rights reserved, also regarding any disposal, exploitation, reproduction, editing, distribution,<br>
as well as in the event of applications for industrial property rights.<br>
*****************************************************************************************************<br>
DESCRIPTION:<br>
Writes a parameter FB's stStaging as the gateway does over ADS (docs/config-contract.md): the version the set is<br>
based on, a stage id, and bStaged (a set, written to stStaged before) or bReset last. ST cannot assign to an FB's<br>
output, so the tests pass the address of vo_Config.stStaging, as ADS writes into the PLC's memory.<br>
*****************************************************************************************************<br>
OUTPUT VALUES:<br>
FALSE for a null pointer.<br>
*****************************************************************************************************<br>
VERSION         ¦ DATE       ¦ NAME      ¦ CHANGE<br>
Syn_Config 2.0.0 ¦ 2026-11-11 ¦ J.Willner ¦ Unit tests<br>
****************************************************************************************************)
FUNCTION _FC_TestConfigStage : BOOL
VAR_INPUT
	vi_p_Staging						: POINTER TO SynConfig.ST_ConfigStaging;	// ADR(fb_Param.vo_Config.stStaging)
	vi_udn_BaseVersion					: UDINT;	// [-] active version the set is based on
	vi_udn_StageId						: UDINT;	// [-] the gateway's id of this staging
	vi_b_Reset							: BOOL;	// [-] TRUE: a reset instead of a staged set
END_VAR

_FC_TestConfigStage := vi_p_Staging <> 0;
IF NOT _FC_TestConfigStage THEN
	RETURN;
END_IF
vi_p_Staging^.bStaged := FALSE;
vi_p_Staging^.nBaseVersion := vi_udn_BaseVersion;
vi_p_Staging^.nStageId := vi_udn_StageId;
vi_p_Staging^.bReset := vi_b_Reset;
vi_p_Staging^.bStaged := NOT vi_b_Reset;

END_FUNCTION

// ---- POUs/Tests/_FB_TestConfigRobot.TcPOU
(****************************************************************************************************<br>
© Syntegon Group.<br>
All rights reserved, also regarding any disposal, exploitation, reproduction, editing, distribution,<br>
as well as in the event of applications for industrial property rights.<br>
*****************************************************************************************************<br>
DESCRIPTION:<br>
TcUnit test suite of the robots' parameter FBs (SynConfig._FB_ConfigDelta, _FB_ConfigXtsGantry,<br>
_FB_ConfigXtsLoop, _FB_ConfigCartesian): which staged sets are rejected and why (zones, gripper fingers, track<br>
modules), and m_PassOn handing the effective values on to the robot's Syn_Visu FB, its config version changing<br>
only when a value does, its lists shrinking with the set.<br>
*****************************************************************************************************<br>
VERSION         ¦ DATE       ¦ NAME      ¦ CHANGE<br>
Syn_Config 2.0.0 ¦ 2026-11-11 ¦ J.Willner ¦ Unit tests<br>
****************************************************************************************************)
FUNCTION_BLOCK _FB_TestConfigRobot EXTENDS TcUnit.FB_TestSuite

m_DeltaRejectsInvalidZonesAndFingers();
m_XtsTracksRejectInvalidModules();
m_CartesianTakesOverFingers();
m_DeltaPassOn();
m_DeltaPassOnShrinksLists();
m_XtsGantryPassOnModules();

(****************************************************************************************************<br>
© Syntegon Group.<br>
All rights reserved, also regarding any disposal, exploitation, reproduction, editing, distribution,<br>
as well as in the event of applications for industrial property rights.<br>
*****************************************************************************************************<br>
DESCRIPTION:<br>
A Cartesian robot's set takes its gripper fingers over with their offsets on the flange (ADR 0018); a finger<br>
without a height is rejected.<br>
****************************************************************************************************)
METHOD PRIVATE m_CartesianTakesOverFingers
VAR_INST
	fb_TempParam						: SynConfig._FB_ConfigCartesian;
	TempDefault							: SynConfig.ST_ConfigCartesianParam;
	TempSet								: SynConfig.ST_ConfigCartesianSet;
	b_TempDone							: BOOL;	// the test ran
END_VAR
VAR
	TempStaged							: SynConfig.ST_ConfigCartesianParam;
	p_TempStaged						: POINTER TO SynConfig.ST_ConfigCartesianParam;
END_VAR
TEST('ConfigCartesianTakesOverFingers');
IF b_TempDone THEN
	RETURN;
END_IF
b_TempDone := TRUE;

p_TempStaged := ADR(fb_TempParam.vo_Config.stStaged);
TempStaged.nFingerCount := 2;
TempStaged.aFingers[0].fDiameter := 30;
TempStaged.aFingers[0].fHeight := 60;
TempStaged.aFingers[1].fDiameter := 30;
TempStaged.aFingers[1].fHeight := 0;
TempStaged.aFingers[1].stOffset.fY := -45;
TempStaged.aFingers[1].stOffset.fRz := 90;

p_TempStaged^ := TempStaged;
_FC_TestConfigStage(vi_p_Staging := ADR(fb_TempParam.vo_Config.stStaging), vi_udn_BaseVersion := 0, vi_udn_StageId := 1,
	vi_b_Reset := FALSE);
AssertFalse(Condition := fb_TempParam.m_Cycle(vio_Default := TempDefault, vio_Set := TempSet, vi_b_ApplyAllowed := TRUE),
	Message := 'finger without a height: not taken over');
AssertEquals_STRING(Expected := 'Finger 2 has no diameter or height', Actual := fb_TempParam.vo_Config.stStatus.sMessage,
	Message := 'reason');

TempStaged.aFingers[1].fHeight := 60;
p_TempStaged^ := TempStaged;
_FC_TestConfigStage(vi_p_Staging := ADR(fb_TempParam.vo_Config.stStaging), vi_udn_BaseVersion := 0, vi_udn_StageId := 2,
	vi_b_Reset := FALSE);
AssertTrue(Condition := fb_TempParam.m_Cycle(vio_Default := TempDefault, vio_Set := TempSet, vi_b_ApplyAllowed := TRUE),
	Message := 'valid fingers taken over');
AssertEquals_UINT(Expected := 2, Actual := fb_TempParam.vo_Config.stActive.nFingerCount, Message := 'two fingers effective');
AssertEquals_LREAL(Expected := -45, Actual := fb_TempParam.vo_Config.stActive.aFingers[1].stOffset.fY, Delta := 0.001,
	Message := 'offset Y kept');
AssertEquals_LREAL(Expected := 90, Actual := fb_TempParam.vo_Config.stActive.aFingers[1].stOffset.fRz, Delta := 0.001,
	Message := 'offset rotation kept');

TEST_FINISHED();
END_METHOD

(****************************************************************************************************<br>
© Syntegon Group.<br>
All rights reserved, also regarding any disposal, exploitation, reproduction, editing, distribution,<br>
as well as in the event of applications for industrial property rights.<br>
*****************************************************************************************************<br>
DESCRIPTION:<br>
m_PassOn hands a Delta's effective pose, origin shift, working area, limit areas, zones and fingers with their offsets<br>
on to its Syn_Visu FB. Called every cycle with the same values, it leaves Syn_Visu's config version alone.<br>
****************************************************************************************************)
METHOD PRIVATE m_DeltaPassOn
VAR_INST
	fb_TempParam						: SynConfig._FB_ConfigDelta;
	fb_TempVisu							: _FB_VisuDelta;
	TempVisuManifest					: ST_VisuManifest;
	TempDefault							: SynConfig.ST_ConfigDeltaParam;
	TempSet								: SynConfig.ST_ConfigDeltaSet;
	b_TempDone							: BOOL;	// the test ran
END_VAR
VAR
	udn_TempVersion						: UDINT;	// [-] Syn_Visu's config version after the first m_PassOn
END_VAR
TEST('ConfigDeltaPassOn');
IF b_TempDone THEN
	RETURN;
END_IF
b_TempDone := TRUE;

fb_TempVisu.m_Register(vio_Manifest := TempVisuManifest, vi_udn_Id := 10, vi_str_Name := 'Delta 1');
TempDefault := m_DeltaSet(vi_un_Zones := 2, vi_un_Fingers := 3);
fb_TempParam.m_Cycle(vio_Default := TempDefault, vio_Set := TempSet, vi_b_ApplyAllowed := TRUE);
AssertTrue(Condition := fb_TempParam.m_PassOn(vio_Visu := fb_TempVisu), Message := 'passed on');

AssertEquals_LREAL(Expected := 1000, Actual := fb_TempVisu.vo_Visu.stConfig.stPose.fX, Delta := 0.001, Message := 'pose X');
AssertEquals_LREAL(Expected := 1900, Actual := fb_TempVisu.vo_Visu.stConfig.stPose.fZ, Delta := 0.001, Message := 'pose Z');

AssertEquals_LREAL(Expected := 20, Actual := fb_TempVisu.vo_Visu.stConfig.stOriginShift.fY, Delta := 0.001,
	Message := 'origin shift');
AssertEquals_LREAL(Expected := 700, Actual := fb_TempVisu.vo_Visu.stConfig.stWorkingArea.fRadius, Delta := 0.001,
	Message := 'working area');
AssertTrue(Condition := fb_TempVisu.vo_Visu.stConfig.stLimitArea.bActive, Message := 'limit area set');
AssertEquals_LREAL(Expected := 400, Actual := fb_TempVisu.vo_Visu.stConfig.stLimitArea.fXMax, Delta := 0.001,
	Message := 'limit area values');
AssertFalse(Condition := fb_TempVisu.vo_Visu.stConfig.stTcpLimitArea.bActive, Message := 'no TCP limit area');
AssertEquals_UINT(Expected := 2, Actual := fb_TempVisu.vo_Visu.stConfig.nZoneCount, Message := 'two zones');
AssertEquals_LREAL(Expected := 2000, Actual := fb_TempVisu.vo_Visu.stConfig.aZones[1].fStart, Delta := 0.001,
	Message := 'zone 2 start');
AssertEquals_UINT(Expected := 3, Actual := fb_TempVisu.vo_Visu.stConfig.nFingerCount, Message := 'three fingers');
AssertEquals_LREAL(Expected := 40, Actual := fb_TempVisu.vo_Visu.stConfig.aFingers[2].fDiameter, Delta := 0.001,
	Message := 'finger 3 diameter');
AssertEquals_LREAL(Expected := 120, Actual := fb_TempVisu.vo_Visu.stConfig.aFingers[2].stOffset.fX, Delta := 0.001,
	Message := 'finger 3 offset X');
AssertEquals_LREAL(Expected := 60, Actual := fb_TempVisu.vo_Visu.stConfig.aFingers[2].stOffset.fRz, Delta := 0.001,
	Message := 'finger 3 offset rotation');

udn_TempVersion := TempVisuManifest.nConfigVersion;
fb_TempParam.m_Cycle(vio_Default := TempDefault, vio_Set := TempSet, vi_b_ApplyAllowed := TRUE);
fb_TempParam.m_PassOn(vio_Visu := fb_TempVisu);
AssertEquals_UDINT(Expected := udn_TempVersion, Actual := TempVisuManifest.nConfigVersion,
	Message := 'same values again: config version unchanged');

TEST_FINISHED();
END_METHOD

(****************************************************************************************************<br>
© Syntegon Group.<br>
All rights reserved, also regarding any disposal, exploitation, reproduction, editing, distribution,<br>
as well as in the event of applications for industrial property rights.<br>
*****************************************************************************************************<br>
DESCRIPTION:<br>
Syn_Visu's zone and finger counts only grow, so m_PassOn clears them when the effective set has fewer: after a<br>
set with fewer zones and no fingers the visualisation has exactly those; an inactive limit area is cleared.<br>
****************************************************************************************************)
METHOD PRIVATE m_DeltaPassOnShrinksLists
VAR_INST
	fb_TempParam						: SynConfig._FB_ConfigDelta;
	fb_TempVisu							: _FB_VisuDelta;
	TempDefault							: SynConfig.ST_ConfigDeltaParam;
	TempSet								: SynConfig.ST_ConfigDeltaSet;
	b_TempDone							: BOOL;	// the test ran
END_VAR
TEST('ConfigDeltaPassOnShrinksLists');
IF b_TempDone THEN
	RETURN;
END_IF
b_TempDone := TRUE;

TempDefault := m_DeltaSet(vi_un_Zones := 3, vi_un_Fingers := 3);
fb_TempParam.m_Cycle(vio_Default := TempDefault, vio_Set := TempSet, vi_b_ApplyAllowed := TRUE);
fb_TempParam.m_PassOn(vio_Visu := fb_TempVisu);
AssertEquals_UINT(Expected := 3, Actual := fb_TempVisu.vo_Visu.stConfig.nZoneCount, Message := 'three zones first');
AssertEquals_UINT(Expected := 3, Actual := fb_TempVisu.vo_Visu.stConfig.nFingerCount, Message := 'three fingers first');

(* The program values change: one zone, no gripper, no limit area. *)
TempDefault := m_DeltaSet(vi_un_Zones := 1, vi_un_Fingers := 0);
TempDefault.stLimitArea.bActive := FALSE;
fb_TempParam.m_Cycle(vio_Default := TempDefault, vio_Set := TempSet, vi_b_ApplyAllowed := TRUE);
fb_TempParam.m_PassOn(vio_Visu := fb_TempVisu);
AssertEquals_UINT(Expected := 1, Actual := fb_TempVisu.vo_Visu.stConfig.nZoneCount, Message := 'one zone left');
AssertEquals_LREAL(Expected := 1000, Actual := fb_TempVisu.vo_Visu.stConfig.aZones[0].fStart, Delta := 0.001,
	Message := 'the remaining zone');
AssertEquals_UINT(Expected := 0, Actual := fb_TempVisu.vo_Visu.stConfig.nFingerCount, Message := 'no fingers left');
AssertFalse(Condition := fb_TempVisu.vo_Visu.stConfig.stLimitArea.bActive, Message := 'limit area cleared');

TEST_FINISHED();
END_METHOD

(****************************************************************************************************<br>
© Syntegon Group.<br>
All rights reserved, also regarding any disposal, exploitation, reproduction, editing, distribution,<br>
as well as in the event of applications for industrial property rights.<br>
*****************************************************************************************************<br>
DESCRIPTION:<br>
A Delta set is rejected with the reason for a zone on no conveyor, a finger without a diameter or height, or more<br>
zones or fingers than the lists hold; zones are checked before fingers. A valid set is then taken over.<br>
****************************************************************************************************)
METHOD PRIVATE m_DeltaRejectsInvalidZonesAndFingers
VAR_INST
	fb_TempParam						: SynConfig._FB_ConfigDelta;
	TempDefault							: SynConfig.ST_ConfigDeltaParam;
	TempSet								: SynConfig.ST_ConfigDeltaSet;
	b_TempDone							: BOOL;	// the test ran
END_VAR
VAR
	TempStaged							: SynConfig.ST_ConfigDeltaParam;
	p_TempStaged						: POINTER TO SynConfig.ST_ConfigDeltaParam;
END_VAR
TEST('ConfigDeltaRejectsInvalidZonesAndFingers');
IF b_TempDone THEN
	RETURN;
END_IF
b_TempDone := TRUE;

TempDefault := m_DeltaSet(vi_un_Zones := 1, vi_un_Fingers := 1);
p_TempStaged := ADR(fb_TempParam.vo_Config.stStaged);

(* A zone on no conveyor, and a finger without a diameter: the zone is named. *)
TempStaged := m_DeltaSet(vi_un_Zones := 2, vi_un_Fingers := 2);
TempStaged.aZones[0].nConveyorId := 0;
TempStaged.aFingers[1].fDiameter := 0;
p_TempStaged^ := TempStaged;
_FC_TestConfigStage(vi_p_Staging := ADR(fb_TempParam.vo_Config.stStaging), vi_udn_BaseVersion := 0, vi_udn_StageId := 1,
	vi_b_Reset := FALSE);
AssertFalse(Condition := fb_TempParam.m_Cycle(vio_Default := TempDefault, vio_Set := TempSet, vi_b_ApplyAllowed := TRUE),
	Message := 'zone on no conveyor: not taken over');
AssertTrue(Condition := fb_TempParam.vo_Config.stStatus.eResult = SynConfig.E_ConfigResult.REJECTED, Message := 'rejected');
AssertEquals_STRING(Expected := 'Zone 1 lies on no conveyor', Actual := fb_TempParam.vo_Config.stStatus.sMessage,
	Message := 'reason: the zone, checked first');

(* A finger without a diameter. *)
TempStaged := m_DeltaSet(vi_un_Zones := 2, vi_un_Fingers := 2);
TempStaged.aFingers[1].fDiameter := 0;
p_TempStaged^ := TempStaged;
_FC_TestConfigStage(vi_p_Staging := ADR(fb_TempParam.vo_Config.stStaging), vi_udn_BaseVersion := 0, vi_udn_StageId := 2,
	vi_b_Reset := FALSE);
fb_TempParam.m_Cycle(vio_Default := TempDefault, vio_Set := TempSet, vi_b_ApplyAllowed := TRUE);
AssertEquals_STRING(Expected := 'Finger 2 has no diameter or height', Actual := fb_TempParam.vo_Config.stStatus.sMessage,
	Message := 'reason: finger without a diameter');

(* A finger without a height. *)
TempStaged := m_DeltaSet(vi_un_Zones := 2, vi_un_Fingers := 2);
TempStaged.aFingers[0].fHeight := 0;
p_TempStaged^ := TempStaged;
_FC_TestConfigStage(vi_p_Staging := ADR(fb_TempParam.vo_Config.stStaging), vi_udn_BaseVersion := 0, vi_udn_StageId := 3,
	vi_b_Reset := FALSE);
fb_TempParam.m_Cycle(vio_Default := TempDefault, vio_Set := TempSet, vi_b_ApplyAllowed := TRUE);
AssertEquals_STRING(Expected := 'Finger 1 has no diameter or height', Actual := fb_TempParam.vo_Config.stStatus.sMessage,
	Message := 'reason: finger without a height');

(* More zones, then more fingers than the lists hold. *)
TempStaged := m_DeltaSet(vi_un_Zones := 2, vi_un_Fingers := 2);
TempStaged.nZoneCount := VISU_GlobalConst_Param.VISU_un_MAX_ZONES + 1;
p_TempStaged^ := TempStaged;
_FC_TestConfigStage(vi_p_Staging := ADR(fb_TempParam.vo_Config.stStaging), vi_udn_BaseVersion := 0, vi_udn_StageId := 4,
	vi_b_Reset := FALSE);
fb_TempParam.m_Cycle(vio_Default := TempDefault, vio_Set := TempSet, vi_b_ApplyAllowed := TRUE);
AssertEquals_STRING(Expected := CONCAT('More than ', CONCAT(UINT_TO_STRING(VISU_GlobalConst_Param.VISU_un_MAX_ZONES), ' zones')),
	Actual := fb_TempParam.vo_Config.stStatus.sMessage, Message := 'reason: too many zones');
TempStaged := m_DeltaSet(vi_un_Zones := 2, vi_un_Fingers := 2);
TempStaged.nFingerCount := VISU_GlobalConst_Param.VISU_un_MAX_FINGERS + 1;
p_TempStaged^ := TempStaged;
_FC_TestConfigStage(vi_p_Staging := ADR(fb_TempParam.vo_Config.stStaging), vi_udn_BaseVersion := 0, vi_udn_StageId := 5,
	vi_b_Reset := FALSE);
fb_TempParam.m_Cycle(vio_Default := TempDefault, vio_Set := TempSet, vi_b_ApplyAllowed := TRUE);
AssertEquals_STRING(Expected := CONCAT('More than ', CONCAT(UINT_TO_STRING(VISU_GlobalConst_Param.VISU_un_MAX_FINGERS), ' fingers')),
	Actual := fb_TempParam.vo_Config.stStatus.sMessage, Message := 'reason: too many fingers');
AssertFalse(Condition := TempSet.bValid, Message := 'no set taken over so far');

(* A valid set. *)
TempStaged := m_DeltaSet(vi_un_Zones := 2, vi_un_Fingers := 2);
p_TempStaged^ := TempStaged;
_FC_TestConfigStage(vi_p_Staging := ADR(fb_TempParam.vo_Config.stStaging), vi_udn_BaseVersion := 0, vi_udn_StageId := 6,
	vi_b_Reset := FALSE);
AssertTrue(Condition := fb_TempParam.m_Cycle(vio_Default := TempDefault, vio_Set := TempSet, vi_b_ApplyAllowed := TRUE),
	Message := 'valid set taken over');
AssertEquals_UINT(Expected := 2, Actual := fb_TempParam.m_ZoneCount(), Message := 'its zones effective');

TEST_FINISHED();
END_METHOD

(****************************************************************************************************<br>
© Syntegon Group.<br>
All rights reserved, also regarding any disposal, exploitation, reproduction, editing, distribution,<br>
as well as in the event of applications for industrial property rights.<br>
*****************************************************************************************************<br>
DESCRIPTION:<br>
A Delta parameter set that can be taken over: origin shift (10, 20, 30), a working area of radius 700, a limit<br>
area, no TCP limit area, vi_un_Zones zones on conveyor 1 (zone n from n * 1000) and vi_un_Fingers fingers of<br>
40 x 50 mm, finger n at X = (n - 1) * 60 mm, turned by (n - 1) * 30 degrees.<br>
****************************************************************************************************)
METHOD PRIVATE m_DeltaSet : SynConfig.ST_ConfigDeltaParam
VAR_INPUT
	vi_un_Zones							: UINT;	// [-] zones, at most VISU_un_MAX_ZONES
	vi_un_Fingers						: UINT;	// [-] fingers, at most VISU_un_MAX_FINGERS
END_VAR
VAR
	un_TempIndex						: UINT;
END_VAR
m_DeltaSet.stPose.fX := 1000;
m_DeltaSet.stPose.fZ := 1900;
m_DeltaSet.stOriginShift.fX := 10;
m_DeltaSet.stOriginShift.fY := 20;
m_DeltaSet.stOriginShift.fZ := 30;
m_DeltaSet.stWorkingArea.fRadius := 700;
m_DeltaSet.stWorkingArea.fZMin := -1300;
m_DeltaSet.stWorkingArea.fZMax := -700;
m_DeltaSet.stLimitArea.fXMin := -500;
m_DeltaSet.stLimitArea.fXMax := 400;
m_DeltaSet.stLimitArea.fYMin := -600;
m_DeltaSet.stLimitArea.fYMax := 600;
m_DeltaSet.stLimitArea.fZMin := -1300;
m_DeltaSet.stLimitArea.fZMax := -700;
m_DeltaSet.stLimitArea.bActive := TRUE;

m_DeltaSet.nZoneCount := MIN(vi_un_Zones, VISU_GlobalConst_Param.VISU_un_MAX_ZONES);
FOR un_TempIndex := 1 TO m_DeltaSet.nZoneCount DO
	m_DeltaSet.aZones[un_TempIndex - 1].nConveyorId := 1;
	m_DeltaSet.aZones[un_TempIndex - 1].fStart := UINT_TO_LREAL(un_TempIndex) * 1000;
	m_DeltaSet.aZones[un_TempIndex - 1].fEnd := UINT_TO_LREAL(un_TempIndex) * 1000 + 500;
END_FOR

m_DeltaSet.nFingerCount := MIN(vi_un_Fingers, VISU_GlobalConst_Param.VISU_un_MAX_FINGERS);
FOR un_TempIndex := 1 TO m_DeltaSet.nFingerCount DO
	m_DeltaSet.aFingers[un_TempIndex - 1].fDiameter := 40;
	m_DeltaSet.aFingers[un_TempIndex - 1].fHeight := 50;
	m_DeltaSet.aFingers[un_TempIndex - 1].stOffset.fX := UINT_TO_LREAL(un_TempIndex - 1) * 60;
	m_DeltaSet.aFingers[un_TempIndex - 1].stOffset.fRz := UINT_TO_LREAL(un_TempIndex - 1) * 30;
END_FOR
END_METHOD

(****************************************************************************************************<br>
© Syntegon Group.<br>
All rights reserved, also regarding any disposal, exploitation, reproduction, editing, distribution,<br>
as well as in the event of applications for industrial property rights.<br>
*****************************************************************************************************<br>
DESCRIPTION:<br>
m_PassOn hands an XTS gantry's effective track modules on to its Syn_Visu FB, leaves the config version alone<br>
while they stay, and shortens the visualisation's track when the set has fewer modules.<br>
****************************************************************************************************)
METHOD PRIVATE m_XtsGantryPassOnModules
VAR_INST
	fb_TempParam						: SynConfig._FB_ConfigXtsGantry;
	fb_TempVisu							: _FB_VisuXtsGantry;
	TempVisuManifest					: ST_VisuManifest;
	TempDefault							: SynConfig.ST_ConfigXtsGantryParam;
	TempSet								: SynConfig.ST_ConfigXtsGantrySet;
	b_TempDone							: BOOL;	// the test ran
END_VAR
VAR
	un_TempIndex						: UINT;
	udn_TempVersion						: UDINT;	// [-] Syn_Visu's config version after the first m_PassOn
END_VAR
TEST('ConfigXtsGantryPassOnModules');
IF b_TempDone THEN
	RETURN;
END_IF
b_TempDone := TRUE;

fb_TempVisu.m_Register(vio_Manifest := TempVisuManifest, vi_udn_Id := 30, vi_str_Name := 'IDH');
TempDefault.nModuleCount := 4;
FOR un_TempIndex := 0 TO 3 DO
	TempDefault.aModules[un_TempIndex].eKind := E_VisuModuleKind.STRAIGHT;
	TempDefault.aModules[un_TempIndex].fLength := 250;
END_FOR
fb_TempParam.m_Cycle(vio_Default := TempDefault, vio_Set := TempSet, vi_b_ApplyAllowed := TRUE);
AssertTrue(Condition := fb_TempParam.m_PassOn(vio_Visu := fb_TempVisu), Message := 'passed on');
AssertEquals_UINT(Expected := 4, Actual := fb_TempVisu.vo_Visu.stConfig.nModuleCount, Message := 'four modules');
AssertEquals_LREAL(Expected := 250, Actual := fb_TempVisu.vo_Visu.stConfig.aModules[3].fLength, Delta := 0.001,
	Message := 'module 4 length');

udn_TempVersion := TempVisuManifest.nConfigVersion;
fb_TempParam.m_PassOn(vio_Visu := fb_TempVisu);
AssertEquals_UDINT(Expected := udn_TempVersion, Actual := TempVisuManifest.nConfigVersion,
	Message := 'same modules again: config version unchanged');

TempDefault.nModuleCount := 2;
fb_TempParam.m_Cycle(vio_Default := TempDefault, vio_Set := TempSet, vi_b_ApplyAllowed := TRUE);
fb_TempParam.m_PassOn(vio_Visu := fb_TempVisu);
AssertEquals_UINT(Expected := 2, Actual := fb_TempVisu.vo_Visu.stConfig.nModuleCount, Message := 'track shortened to two modules');

TEST_FINISHED();
END_METHOD

(****************************************************************************************************<br>
© Syntegon Group.<br>
All rights reserved, also regarding any disposal, exploitation, reproduction, editing, distribution,<br>
as well as in the event of applications for industrial property rights.<br>
*****************************************************************************************************<br>
DESCRIPTION:<br>
An XTS gantry or loop set is rejected with the reason for a track without modules, a module without a length or<br>
more modules than the list holds; modules are checked before zones. A valid loop set is then taken over.<br>
****************************************************************************************************)
METHOD PRIVATE m_XtsTracksRejectInvalidModules
VAR_INST
	fb_TempGantryParam					: SynConfig._FB_ConfigXtsGantry;
	fb_TempLoopParam					: SynConfig._FB_ConfigXtsLoop;
	TempGantryDefault					: SynConfig.ST_ConfigXtsGantryParam;
	TempGantrySet						: SynConfig.ST_ConfigXtsGantrySet;
	TempLoopDefault						: SynConfig.ST_ConfigXtsLoopParam;
	TempLoopSet							: SynConfig.ST_ConfigXtsLoopSet;
	b_TempDone							: BOOL;	// the test ran
END_VAR
VAR
	TempGantryStaged					: SynConfig.ST_ConfigXtsGantryParam;
	TempLoopStaged						: SynConfig.ST_ConfigXtsLoopParam;
	p_TempGantryStaged					: POINTER TO SynConfig.ST_ConfigXtsGantryParam;
	p_TempLoopStaged					: POINTER TO SynConfig.ST_ConfigXtsLoopParam;
END_VAR
TEST('ConfigXtsTracksRejectInvalidModules');
IF b_TempDone THEN
	RETURN;
END_IF
b_TempDone := TRUE;

p_TempGantryStaged := ADR(fb_TempGantryParam.vo_Config.stStaged);
p_TempLoopStaged := ADR(fb_TempLoopParam.vo_Config.stStaged);

(* Gantry: a track without modules, also with a zone on no conveyor: the track is named. *)
TempGantryStaged.nModuleCount := 0;
TempGantryStaged.nZoneCount := 1;
TempGantryStaged.aZones[0].nConveyorId := 0;
p_TempGantryStaged^ := TempGantryStaged;
_FC_TestConfigStage(vi_p_Staging := ADR(fb_TempGantryParam.vo_Config.stStaging), vi_udn_BaseVersion := 0, vi_udn_StageId := 1,
	vi_b_Reset := FALSE);
AssertFalse(Condition := fb_TempGantryParam.m_Cycle(vio_Default := TempGantryDefault, vio_Set := TempGantrySet,
	vi_b_ApplyAllowed := TRUE), Message := 'gantry without modules: not taken over');
AssertEquals_STRING(Expected := 'A track without modules', Actual := fb_TempGantryParam.vo_Config.stStatus.sMessage,
	Message := 'reason: no modules, checked first');

(* Gantry: more modules than the list holds. *)
TempGantryStaged.nModuleCount := VISU_GlobalConst_Param.VISU_un_MAX_MODULES + 1;
p_TempGantryStaged^ := TempGantryStaged;
_FC_TestConfigStage(vi_p_Staging := ADR(fb_TempGantryParam.vo_Config.stStaging), vi_udn_BaseVersion := 0, vi_udn_StageId := 2,
	vi_b_Reset := FALSE);
fb_TempGantryParam.m_Cycle(vio_Default := TempGantryDefault, vio_Set := TempGantrySet, vi_b_ApplyAllowed := TRUE);
AssertEquals_STRING(Expected := CONCAT('More than ', CONCAT(UINT_TO_STRING(VISU_GlobalConst_Param.VISU_un_MAX_MODULES),
	' track modules')), Actual := fb_TempGantryParam.vo_Config.stStatus.sMessage, Message := 'reason: too many modules');

(* Loop: module 2 without a length. *)
TempLoopStaged.nModuleCount := 3;
TempLoopStaged.aModules[0].eKind := E_VisuModuleKind.STRAIGHT;
TempLoopStaged.aModules[0].fLength := 250;
TempLoopStaged.aModules[1].eKind := E_VisuModuleKind.CURVE_LEFT;
TempLoopStaged.aModules[1].fLength := 0;
TempLoopStaged.aModules[2].eKind := E_VisuModuleKind.STRAIGHT;
TempLoopStaged.aModules[2].fLength := 250;
p_TempLoopStaged^ := TempLoopStaged;
_FC_TestConfigStage(vi_p_Staging := ADR(fb_TempLoopParam.vo_Config.stStaging), vi_udn_BaseVersion := 0, vi_udn_StageId := 1,
	vi_b_Reset := FALSE);
AssertFalse(Condition := fb_TempLoopParam.m_Cycle(vio_Default := TempLoopDefault, vio_Set := TempLoopSet,
	vi_b_ApplyAllowed := TRUE), Message := 'loop with a module without a length: not taken over');
AssertEquals_STRING(Expected := 'Track module 2 has no length', Actual := fb_TempLoopParam.vo_Config.stStatus.sMessage,
	Message := 'reason: module without a length');

(* Loop: a valid track. *)
TempLoopStaged.aModules[1].fLength := 250;
p_TempLoopStaged^ := TempLoopStaged;
_FC_TestConfigStage(vi_p_Staging := ADR(fb_TempLoopParam.vo_Config.stStaging), vi_udn_BaseVersion := 0, vi_udn_StageId := 2,
	vi_b_Reset := FALSE);
AssertTrue(Condition := fb_TempLoopParam.m_Cycle(vio_Default := TempLoopDefault, vio_Set := TempLoopSet,
	vi_b_ApplyAllowed := TRUE), Message := 'valid loop taken over');
AssertEquals_UINT(Expected := 3, Actual := fb_TempLoopParam.vo_Config.stActive.nModuleCount, Message := 'its modules effective');
AssertTrue(Condition := fb_TempLoopParam.vo_Config.stActive.aModules[1].eKind = E_VisuModuleKind.CURVE_LEFT,
	Message := 'module kind kept');

TEST_FINISHED();
END_METHOD

END_FUNCTION_BLOCK

// ---- POUs/Tests/_FB_TestConfigBodyComponent.TcPOU
(****************************************************************************************************<br>
© Syntegon Group.<br>
All rights reserved, also regarding any disposal, exploitation, reproduction, editing, distribution,<br>
as well as in the event of applications for industrial property rights.<br>
*****************************************************************************************************<br>
DESCRIPTION:<br>
TcUnit test suite of the parameter FBs of components drawn from their bodies (SynConfig._FB_ConfigVision,<br>
_FB_ConfigSensor, _FB_ConfigStation on _FB_ConfigBodyComponent): the component type each registers, a set with<br>
zones taken over and passed on to the Syn_Visu FB, and a zone on no conveyor rejected.<br>
*****************************************************************************************************<br>
VERSION         ¦ DATE       ¦ NAME      ¦ CHANGE<br>
Syn_Config 2.0.0 ¦ 2026-11-11 ¦ J.Willner ¦ Unit tests<br>
****************************************************************************************************)
FUNCTION_BLOCK _FB_TestConfigBodyComponent EXTENDS TcUnit.FB_TestSuite

m_RegisterComponentTypes();
m_VisionZonesTakenOverAndPassedOn();
m_SensorRejectsZoneOnNoConveyor();

(****************************************************************************************************<br>
© Syntegon Group.<br>
All rights reserved, also regarding any disposal, exploitation, reproduction, editing, distribution,<br>
as well as in the event of applications for industrial property rights.<br>
*****************************************************************************************************<br>
DESCRIPTION:<br>
Vision system, product sensor and station share one structure, but each registers its own component type, from<br>
which the gateway knows the component.<br>
****************************************************************************************************)
METHOD PRIVATE m_RegisterComponentTypes
VAR_INST
	fb_TempVisionParam					: SynConfig._FB_ConfigVision;
	fb_TempSensorParam					: SynConfig._FB_ConfigSensor;
	fb_TempStationParam					: SynConfig._FB_ConfigStation;
	TempManifest						: SynConfig.ST_ConfigManifest;
	b_TempDone							: BOOL;	// the test ran
END_VAR
TEST('ConfigRegisterComponentTypes');
IF b_TempDone THEN
	RETURN;
END_IF
b_TempDone := TRUE;

AssertTrue(Condition := fb_TempVisionParam.m_Register(vio_Manifest := TempManifest, vi_udn_Id := 60), Message := 'vision registered');
AssertTrue(Condition := fb_TempSensorParam.m_Register(vio_Manifest := TempManifest, vi_udn_Id := 61), Message := 'sensor registered');
AssertTrue(Condition := fb_TempStationParam.m_Register(vio_Manifest := TempManifest, vi_udn_Id := 70),
	Message := 'station registered');
AssertEquals_UINT(Expected := 3, Actual := TempManifest.nCount, Message := 'three entries');
AssertTrue(Condition := TempManifest.aEntries[0].eType = E_VisuComponentType.VISION, Message := 'vision type');
AssertTrue(Condition := TempManifest.aEntries[1].eType = E_VisuComponentType.SENSOR, Message := 'sensor type');
AssertTrue(Condition := TempManifest.aEntries[2].eType = E_VisuComponentType.STATION, Message := 'station type');

TEST_FINISHED();
END_METHOD

(****************************************************************************************************<br>
© Syntegon Group.<br>
All rights reserved, also regarding any disposal, exploitation, reproduction, editing, distribution,<br>
as well as in the event of applications for industrial property rights.<br>
*****************************************************************************************************<br>
DESCRIPTION:<br>
A product sensor's set with a zone on no conveyor is rejected with the reason; the program values stay.<br>
****************************************************************************************************)
METHOD PRIVATE m_SensorRejectsZoneOnNoConveyor
VAR_INST
	fb_TempParam						: SynConfig._FB_ConfigSensor;
	TempDefault							: SynConfig.ST_ConfigBodyComponentParam;
	TempSet								: SynConfig.ST_ConfigBodyComponentSet;
	b_TempDone							: BOOL;	// the test ran
END_VAR
VAR
	TempStaged							: SynConfig.ST_ConfigBodyComponentParam;
	p_TempStaged						: POINTER TO SynConfig.ST_ConfigBodyComponentParam;
END_VAR
TEST('ConfigSensorRejectsZoneOnNoConveyor');
IF b_TempDone THEN
	RETURN;
END_IF
b_TempDone := TRUE;

TempDefault.stPose.fX := 200;
TempStaged.stPose.fX := 900;
TempStaged.nZoneCount := 2;
TempStaged.aZones[0].nConveyorId := 1;
TempStaged.aZones[1].nConveyorId := 0;
p_TempStaged := ADR(fb_TempParam.vo_Config.stStaged);
p_TempStaged^ := TempStaged;
_FC_TestConfigStage(vi_p_Staging := ADR(fb_TempParam.vo_Config.stStaging), vi_udn_BaseVersion := 0, vi_udn_StageId := 4,
	vi_b_Reset := FALSE);

AssertFalse(Condition := fb_TempParam.m_Cycle(vio_Default := TempDefault, vio_Set := TempSet, vi_b_ApplyAllowed := TRUE),
	Message := 'not taken over');
AssertTrue(Condition := fb_TempParam.vo_Config.stStatus.eResult = SynConfig.E_ConfigResult.REJECTED, Message := 'rejected');
AssertEquals_STRING(Expected := 'Zone 2 lies on no conveyor', Actual := fb_TempParam.vo_Config.stStatus.sMessage, Message := 'reason');
AssertEquals_LREAL(Expected := 200, Actual := fb_TempParam.vo_Config.stActive.stPose.fX, Delta := 0.001,
	Message := 'program values still effective');

TEST_FINISHED();
END_METHOD

(****************************************************************************************************<br>
© Syntegon Group.<br>
All rights reserved, also regarding any disposal, exploitation, reproduction, editing, distribution,<br>
as well as in the event of applications for industrial property rights.<br>
*****************************************************************************************************<br>
DESCRIPTION:<br>
A vision system's staged set with a pose, an origin shift and two zones is taken over; m_Pose gives the pose and<br>
m_PassOn hands pose, origin shift and zones on to the Syn_Visu FB.<br>
****************************************************************************************************)
METHOD PRIVATE m_VisionZonesTakenOverAndPassedOn
VAR_INST
	fb_TempParam						: SynConfig._FB_ConfigVision;
	fb_TempVisu							: _FB_VisuVision;
	TempDefault							: SynConfig.ST_ConfigBodyComponentParam;
	TempSet								: SynConfig.ST_ConfigBodyComponentSet;
	b_TempDone							: BOOL;	// the test ran
END_VAR
VAR
	TempStaged							: SynConfig.ST_ConfigBodyComponentParam;
	p_TempStaged						: POINTER TO SynConfig.ST_ConfigBodyComponentParam;
	TempPose							: ST_VisuPose;
END_VAR
TEST('ConfigVisionZonesTakenOverAndPassedOn');
IF b_TempDone THEN
	RETURN;
END_IF
b_TempDone := TRUE;

TempStaged.stPose.fX := 1500;
TempStaged.stPose.fZ := 1600;
TempStaged.stOriginShift.fZ := -800;
TempStaged.nZoneCount := 2;
TempStaged.aZones[0].nConveyorId := 1;
TempStaged.aZones[0].fStart := 800;
TempStaged.aZones[0].fEnd := 1200;
TempStaged.aZones[1].nConveyorId := 2;
TempStaged.aZones[1].fStart := 300;
TempStaged.aZones[1].fEnd := 300;
p_TempStaged := ADR(fb_TempParam.vo_Config.stStaged);
p_TempStaged^ := TempStaged;
_FC_TestConfigStage(vi_p_Staging := ADR(fb_TempParam.vo_Config.stStaging), vi_udn_BaseVersion := 0, vi_udn_StageId := 1,
	vi_b_Reset := FALSE);

AssertTrue(Condition := fb_TempParam.m_Cycle(vio_Default := TempDefault, vio_Set := TempSet, vi_b_ApplyAllowed := TRUE),
	Message := 'set taken over');
AssertTrue(Condition := fb_TempParam.vo_Config.stStatus.eResult = SynConfig.E_ConfigResult.APPLIED, Message := 'applied');
TempPose := fb_TempParam.m_Pose();
AssertEquals_LREAL(Expected := 1500, Actual := TempPose.fX, Delta := 0.001, Message := 'staged pose effective');

AssertTrue(Condition := fb_TempParam.m_PassOn(vio_Visu := fb_TempVisu), Message := 'passed on');
AssertEquals_LREAL(Expected := 1500, Actual := fb_TempVisu.vo_Visu.stConfig.stPose.fX, Delta := 0.001, Message := 'pose');
AssertEquals_LREAL(Expected := -800, Actual := fb_TempVisu.vo_Visu.stConfig.stOriginShift.fZ, Delta := 0.001,
	Message := 'origin shift');
AssertEquals_UINT(Expected := 2, Actual := fb_TempVisu.vo_Visu.stConfig.nZoneCount, Message := 'two zones');
AssertEquals_UDINT(Expected := 2, Actual := fb_TempVisu.vo_Visu.stConfig.aZones[1].nConveyorId, Message := 'zone 2 conveyor');
AssertEquals_LREAL(Expected := 1200, Actual := fb_TempVisu.vo_Visu.stConfig.aZones[0].fEnd, Delta := 0.001,
	Message := 'zone 1 end');

TEST_FINISHED();
END_METHOD

END_FUNCTION_BLOCK

// ---- POUs/Tests/_FB_TestConfigMachine.TcPOU
(****************************************************************************************************<br>
© Syntegon Group.<br>
All rights reserved, also regarding any disposal, exploitation, reproduction, editing, distribution,<br>
as well as in the event of applications for industrial property rights.<br>
*****************************************************************************************************<br>
DESCRIPTION:<br>
TcUnit test suite of _FB_ConfigMachine: registration with id 0, recipe fields and their program values, a staged<br>
recipe taken over or rejected, a reset, machine commands answered by the application, and the fields' labels,<br>
descriptions and visibility conditions. The tests write<br>
vo_Config through its address, as the gateway writes over ADS.<br>
*****************************************************************************************************<br>
VERSION         ¦ DATE       ¦ NAME      ¦ CHANGE<br>
Syn_Config 2.1.0 ¦ 2026-11-14 ¦ J.Willner ¦ Unit tests of the machine FB (config protocol 3)<br>
Syn_Config 2.2.0 ¦ 2026-11-14 ¦ J.Willner ¦ Labels, descriptions and visibility conditions (protocol 4, #49)<br>
****************************************************************************************************)
FUNCTION_BLOCK _FB_TestConfigMachine EXTENDS TcUnit.FB_TestSuite
VAR
END_VAR

m_RegisterWithIdZero();
m_ProgramValues();
m_RecipeTakenOverAndReset();
m_RecipeRejected();
m_CommandAnswered();
m_TextAndCondition();

(****************************************************************************************************<br>
© Syntegon Group.<br>
All rights reserved, also regarding any disposal, exploitation, reproduction, editing, distribution,<br>
as well as in the event of applications for industrial property rights.<br>
*****************************************************************************************************<br>
DESCRIPTION:<br>
A requested command waits for the application; its answer names the command id, accepted or rejected with the<br>
reason, and the command no longer waits. Without a request nothing can be answered.<br>
****************************************************************************************************)
METHOD PRIVATE m_CommandAnswered
VAR_INST
	fb_TempMachine						: SynConfig._FB_ConfigMachine;
	b_TempDone							: BOOL;	// the test ran
END_VAR
VAR
	p_TempConfig						: POINTER TO SynConfig.ST_ConfigMachine;
END_VAR
TEST('ConfigMachineCommandAnswered');
IF b_TempDone THEN
	RETURN;
END_IF
b_TempDone := TRUE;

AssertTrue(Condition := fb_TempMachine.m_Command() = SynConfig.E_ConfigCommand.NONE, Message := 'nothing waits');
AssertFalse(Condition := fb_TempMachine.m_AnswerCommand(vi_b_Accepted := TRUE, vi_str_Reason := ''), Message := 'nothing to answer');

p_TempConfig := ADR(fb_TempMachine.vo_Config);
p_TempConfig^.stCommand.nCommandId := 7;
p_TempConfig^.stCommand.eCommand := SynConfig.E_ConfigCommand.START;
p_TempConfig^.stCommand.bRequested := TRUE;
AssertTrue(Condition := fb_TempMachine.m_Command() = SynConfig.E_ConfigCommand.START, Message := 'START waits');
AssertTrue(Condition := fb_TempMachine.m_AnswerCommand(vi_b_Accepted := FALSE, vi_str_Reason := 'Not stopped'), Message := 'answered');
AssertEquals_UDINT(Expected := 7, Actual := fb_TempMachine.vo_Config.stCommandStatus.nHandledCommandId, Message := 'command 7 handled');
AssertTrue(Condition := fb_TempMachine.vo_Config.stCommandStatus.eResult = SynConfig.E_ConfigCommandResult.REJECTED, Message := 'rejected');
AssertEquals_STRING(Expected := 'Not stopped', Actual := fb_TempMachine.vo_Config.stCommandStatus.sMessage, Message := 'its reason');
AssertTrue(Condition := fb_TempMachine.m_Command() = SynConfig.E_ConfigCommand.NONE, Message := 'no longer waits');

TEST_FINISHED();
END_METHOD

(****************************************************************************************************<br>
© Syntegon Group.<br>
All rights reserved, also regarding any disposal, exploitation, reproduction, editing, distribution,<br>
as well as in the event of applications for industrial property rights.<br>
*****************************************************************************************************<br>
DESCRIPTION:<br>
The recipe the tests declare: 1 BeltSpeed (NUMBER 0..500, 150), 2 Picks (INTEGER 1..4, 2), 3 Feed (SWITCH, on),<br>
4 Pattern (CHOICE Lanes, Random; 0).<br>
****************************************************************************************************)
METHOD PRIVATE m_DeclareFields
VAR_IN_OUT
	vio_Machine							: SynConfig._FB_ConfigMachine;
END_VAR
vio_Machine.m_DeclareField(vi_un_Field := 1, vi_str_Name := 'BeltSpeed', vi_udn_Group := 1,
	vi_e_Type := SynConfig.E_ConfigFieldType.NUMBER, vi_str_Unit := 'mm/s', vi_lr_Min := 0, vi_lr_Max := 500,
	vi_lr_ProgramValue := 150);
vio_Machine.m_DeclareField(vi_un_Field := 2, vi_str_Name := 'Picks', vi_udn_Group := 0,
	vi_e_Type := SynConfig.E_ConfigFieldType.INTEGER, vi_str_Unit := '', vi_lr_Min := 1, vi_lr_Max := 4,
	vi_lr_ProgramValue := 2);
vio_Machine.m_DeclareField(vi_un_Field := 3, vi_str_Name := 'Feed', vi_udn_Group := 0,
	vi_e_Type := SynConfig.E_ConfigFieldType.SWITCH, vi_str_Unit := '', vi_lr_Min := 0, vi_lr_Max := 0,
	vi_lr_ProgramValue := 1);
vio_Machine.m_DeclareField(vi_un_Field := 4, vi_str_Name := 'Pattern', vi_udn_Group := 0,
	vi_e_Type := SynConfig.E_ConfigFieldType.CHOICE, vi_str_Unit := '', vi_lr_Min := 0, vi_lr_Max := 0,
	vi_lr_ProgramValue := 0);
vio_Machine.m_SetChoice(vi_un_Field := 4, vi_un_Value := 0, vi_str_Text := 'Lanes');
vio_Machine.m_SetChoice(vi_un_Field := 4, vi_un_Value := 1, vi_str_Text := 'Random');
END_METHOD

(****************************************************************************************************<br>
© Syntegon Group.<br>
All rights reserved, also regarding any disposal, exploitation, reproduction, editing, distribution,<br>
as well as in the event of applications for industrial property rights.<br>
*****************************************************************************************************<br>
DESCRIPTION:<br>
Declared fields are listed with their choices; without a recipe the program values apply, typed by m_Value,<br>
m_Integer and m_Switch. A field 0 is refused, an undeclared one gives 0.<br>
****************************************************************************************************)
METHOD PRIVATE m_ProgramValues
VAR_INST
	fb_TempMachine						: SynConfig._FB_ConfigMachine;
	TempSet								: SynConfig.ST_ConfigRecipeSet;
	b_TempDone							: BOOL;	// the test ran
END_VAR
TEST('ConfigMachineProgramValues');
IF b_TempDone THEN
	RETURN;
END_IF
b_TempDone := TRUE;

